       30: // ---- ukonceni handshake: shodit Execute, pockat az kamera shodi stav ----
           "COG_ETIKETA_is3800-ExecuteCommand/JobLoad" := FALSE;
           IF NOT "COG_ETIKETA_is3800-CommandCompleted"
               AND NOT "COG_ETIKETA_is3800-CommandFailed" THEN
               #Kam_Etiketa_Job.krok := 0;
           END_IF;

       ELSE
           #Kam_Etiketa_Job.krok := 0;
   END_CASE;

   // casovac timeoutu bezi v krocich 10..30
   #TIMER.TIMER_3.TON(IN := #Kam_Etiketa_Job.krok >= 10,
                      PT := #Kam_Etiketa_Job.timeout);
   IF #TIMER.TIMER_3.Q AND #Kam_Etiketa_Job.krok = 30 THEN
       #Kam_Etiketa_Job.krok := 0;                         // pojistka, kdyby kamera stav neshodila
   END_IF;

   #Kam_Etiketa_Job.odesli_pamet := "DB_HMI_recype".ODESLI_dATA;

   // kontrola: v klidu musi job v kamere odpovidat recepture
   #Kam_Etiketa_Job.nesouhlasi := #Kam_Etiketa_Job.krok = 0
   AND #Kam_Etiketa_Job.pozadovany > 0
   AND "COG_ETIKETA_is3800-Online"
   AND WORD_TO_INT("COG_ETIKETA_is3800-Current Job ID") <> #Kam_Etiketa_Job.pozadovany;
END_REGION

REGION Network 23: EXTERNAL_TRIGER
   RUNG wire#powerrail
      { S7_Templates := "SrcType := Int" } EQ_Contact(in1 := #SQCR, in2 := #STEP_5_HOME)
      Contact( "INICIALIZACE_RUN" )
      I_Contact( #TRIG.inicial_ok_op )
      Contact( "AUTOMAT" )
      S_Coil( #HMI.reset_fronty )
      S_Coil( #TRIG.inicial_ok_op )
   END_RUNG
   RUNG wire#powerrail
      Contact( "FirstScan" )
      S_Coil( #HMI.reset_fronty )
      Move(in := 0, out1 => "DB_HMI_recype".obsazenost_fronty, out2 => #zpracovani_dat[1].balik_den)
   END_RUNG
   // the same network as SCL:
   IF (#SQCR = #STEP_5_HOME) AND "INICIALIZACE_RUN" AND NOT #TRIG.inicial_ok_op AND "AUTOMAT" THEN
       #HMI.reset_fronty := TRUE;
       #TRIG.inicial_ok_op := TRUE;
   END_IF;
   IF "FirstScan" THEN
       #HMI.reset_fronty := TRUE;
       "DB_HMI_recype".obsazenost_fronty := 0;
       #zpracovani_dat[1].balik_den := 0;
   END_IF;
END_REGION

REGION Network 24: ETERNAL_TRIGR_INICIAL
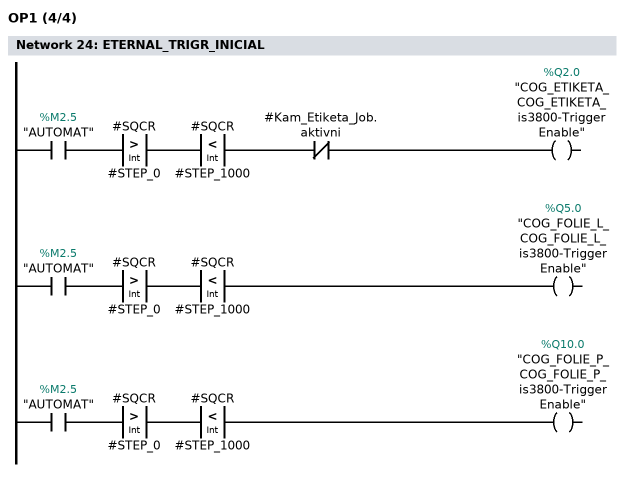
   RUNG wire#powerrail
      Contact( "AUTOMAT" )
      { S7_Templates := "SrcType := Int" } GT_Contact(in1 := #SQCR, in2 := #STEP_0)
      { S7_Templates := "SrcType := Int" } LT_Contact(in1 := #SQCR, in2 := #STEP_1000)
      I_Contact( #Kam_Etiketa_Job.aktivni )
      Coil( "COG_ETIKETA_COG_ETIKETA_is3800-TriggerEnable" )
   END_RUNG
   RUNG wire#powerrail
      Contact( "AUTOMAT" )
      { S7_Templates := "SrcType := Int" } GT_Contact(in1 := #SQCR, in2 := #STEP_0)
      { S7_Templates := "SrcType := Int" } LT_Contact(in1 := #SQCR, in2 := #STEP_1000)
      Coil( "COG_FOLIE_L_COG_FOLIE_L_is3800-TriggerEnable" )
   END_RUNG
   RUNG wire#powerrail
      Contact( "AUTOMAT" )
      { S7_Templates := "SrcType := Int" } GT_Contact(in1 := #SQCR, in2 := #STEP_0)
      { S7_Templates := "SrcType := Int" } LT_Contact(in1 := #SQCR, in2 := #STEP_1000)
      Coil( "COG_FOLIE_P_COG_FOLIE_P_is3800-TriggerEnable" )
   END_RUNG
   // the same network as SCL:
   "COG_ETIKETA_COG_ETIKETA_is3800-TriggerEnable" := "AUTOMAT" AND (#SQCR > #STEP_0) AND (#SQCR < #STEP_1000) AND NOT #Kam_Etiketa_Job.aktivni;
   "COG_FOLIE_L_COG_FOLIE_L_is3800-TriggerEnable" := "AUTOMAT" AND (#SQCR > #STEP_0) AND (#SQCR < #STEP_1000);
   "COG_FOLIE_P_COG_FOLIE_P_is3800-TriggerEnable" := "AUTOMAT" AND (#SQCR > #STEP_0) AND (#SQCR < #STEP_1000);
END_REGION

REGION Network 25: hmi
END_REGION

REGION Network 26 (SCL): VYRAZENI MANUAL
   (* #Test_tp_ka12(IN := "DB_Manual".test_vyr,
                 PT := T#500MS);

   "-KA12" := #Test_tp_ka12.Q;

   // testovací bit se sám shodí → každý Modify TRUE = jeden pulz
   IF "DB_Manual".test_vyr THEN
       "DB_Manual".test_vyr := FALSE;
   END_IF; *)
END_REGION
END_FUNCTION_BLOCK

FUNCTION_BLOCK "FB_CamManual"
{ S7_Optimized_Access := 'TRUE' }
VERSION : 0.1
   VAR_INPUT 
      xManEtiketa : Bool;   // ruční test etiketa
      xManFolie : Bool;   // ruční test folie
      tLightDelay : Time := T#100ms;   // náběh světel
      tTrigPulse : Time := T#50ms;   // d0lka triggeru
   END_VAR

   VAR 
      tonEt {InstructionName := 'TON_TIME'; LibVersion := '1.0'; S7_SetPoint := 'False'} : TON_TIME;
      tpEt {InstructionName := 'TP_TIME'; LibVersion := '1.0'} : TP_TIME;
      tonFo {InstructionName := 'TON_TIME'; LibVersion := '1.0'} : TON_TIME;
      tpFo {InstructionName := 'TP_TIME'; LibVersion := '1.0'} : TP_TIME;
   END_VAR


BEGIN
	// ---------- ETIKETA ----------
	#tonEt(IN := #xManEtiketa,
	       PT := #tLightDelay);
	#tpEt(IN := #tonEt.Q,
	      PT := #tTrigPulse);
	
	IF #xManEtiketa THEN
	    "-KA1" := TRUE;
	    "-KA2" := TRUE;
	END_IF;
	IF #tpEt.Q THEN
	    "COG_ETIKETA_COG_ETIKETA_is3800-Trigger" := TRUE;
	END_IF;
	
	// ---------- FÓLIE ----------
	#tonFo(IN := #xManFolie,
	       PT := #tLightDelay);
	#tpFo(IN := #tonFo.Q,
	      PT := #tTrigPulse);
	
	IF #xManFolie THEN
	    "-KA3" := TRUE;
	    "-KA4" := TRUE;
	    "-KA5" := TRUE;
	END_IF;
	IF #tpFo.Q THEN
	    "COG_FOLIE_L_is3800-Trigger" := TRUE;
	    "COG_FOLIE_P_is3800-Trigger" := TRUE;
	END_IF;
END_FUNCTION_BLOCK

FUNCTION_BLOCK "OP2"   // FB51, LAD
{ S7_Optimized_Access := 'FALSE' }
// stored: AutoNumber false, SetENOAutomatically false
   VAR
      CONTROL_MAN : Struct
         B0 : Bool;
         B1 : Bool;
         B2 : Bool;
         B3 : Bool;
         B4 : Bool;
         B5 : Bool;
         B6 : Bool;
         B7 : Bool;
         B8 : Bool;
         B9 : Bool;
         odfuk_1 : Bool;
         odfuk_2 : Bool;
         B12 : Bool;
         B13 : Bool;
         B14 : Bool;
         B15 : Bool;
         B16 : Bool;
         B17 : Bool;
         B18 : Bool;
         B19 : Bool;
         B20 : Bool;
         B21 : Bool;
         B22 : Bool;
         B23 : Bool;
         B24 : Bool;
         B25 : Bool;
         B26 : Bool;
         B27 : Bool;
         B28 : Bool;
         B29 : Bool;
         B30 : Bool;
         B31 : Bool;
      END_STRUCT;
      CONTROL_AUTOMAT : Struct
         connect : Bool;
         send : Bool;
         reciv : Bool;
         trcv : Bool;
         discon : Bool;
         B5 : Bool;
         B6 : Bool;
         B7 : Bool;
         B8 : Bool;
         B9 : Bool;
         B10 : Bool;
         B11 : Bool;
         B12 : Bool;
         B13 : Bool;
         B14 : Bool;
         B15 : Bool;
         B16 : Bool;
         B17 : Bool;
         B18 : Bool;
         B19 : Bool;
         B20 : Bool;
         B21 : Bool;
         B22 : Bool;
         B23 : Bool;
         B24 : Bool;
         B25 : Bool;
         B26 : Bool;
         B27 : Bool;
         B28 : Bool;
         B29 : Bool;
         B30 : Bool;
         B31 : Bool;
      END_STRUCT;
      SENSORS : Struct
         S0 : Bool;
         S1 : Bool;
         S2 : Bool;
         S3 : Bool;
         S4 : Bool;
         S5 : Bool;
         S6 : Bool;
         S7 : Bool;
         S8 : Bool;   // KARUSEL JE NATOČEN PŘÍPRAVKEM A K BRÁNĚ
         S9 : Bool;
         S10 : Bool;
         S11 : Bool;
         S12 : Bool;
         S13 : Bool;
         S14 : Bool;
         S15 : Bool;
         S16 : Bool;
         S17 : Bool;
         S18 : Bool;
         S19 : Bool;
         S20 : Bool;
         S21 : Bool;
         S22 : Bool;
         S23 : Bool;
         S24 : Bool;
         S25 : Bool;
         S26 : Bool;
         S27 : Bool;
         S28 : Bool;
         S29 : Bool;
         S30 : Bool;
         S31 : Bool;
      END_STRUCT;
      SENSORS_1 : Struct
         S0 : Bool;
         S1 : Bool;
         S2 : Bool;
         S3 : Bool;
         S4 : Bool;
         S5 : Bool;
         S6 : Bool;
         S7 : Bool;
         S8 : Bool;
         S9 : Bool;
         S10 : Bool;
         S11 : Bool;
         S12 : Bool;
         S13 : Bool;
         S14 : Bool;
         S15 : Bool;
         S16 : Bool;
         S17 : Bool;
         S18 : Bool;
         S19 : Bool;
         S20 : Bool;
         S21 : Bool;
         S22 : Bool;
         S23 : Bool;
         S24 : Bool;
         S25 : Bool;
         S26 : Bool;
         S27 : Bool;
         S28 : Bool;
         S29 : Bool;
         S30 : Bool;
         S31 : Bool;
      END_STRUCT;
      S_0 : "SENSOR";
      S_1 : "SENSOR";
      S_2 { S7_SetPoint := 'True'} : "SENSOR";
      S_3 { S7_SetPoint := 'True'} : "SENSOR";
      S_4 { S7_SetPoint := 'True'} : "SENSOR";
      S_5 { S7_SetPoint := 'True'} : "SENSOR";
      S_6 { S7_SetPoint := 'True'} : "SENSOR";
      S_7 { S7_SetPoint := 'True'} : "SENSOR";
      S_8 { S7_SetPoint := 'True'} : "SENSOR";
      S_9 { S7_SetPoint := 'True'} : "SENSOR";
      S_10 { S7_SetPoint := 'True'} : "SENSOR";
      S_11 { S7_SetPoint := 'True'} : "SENSOR";
      S_12 { S7_SetPoint := 'True'} : "SENSOR";
      S_13 { S7_SetPoint := 'True'} : "SENSOR";
      S_14 { S7_SetPoint := 'True'} : "SENSOR";
      S_15 { S7_SetPoint := 'True'} : "SENSOR";
      S_16 { S7_SetPoint := 'True'} : "SENSOR";
      M_1 : "MOTOR_CONTROL_BLOCK";
      M_2 { S7_SetPoint := 'True'} : "MOTOR_CONTROL_BLOCK";
      M_3 { S7_SetPoint := 'True'} : "MOTOR_CONTROL_BLOCK";
      SQCR { S7_SetPoint := 'True'} : Int;
      hmi_sqcr : Int;
      TRIG : Struct
         inicial_ok_op : Bool;
         T2 : Bool;
         T3 : Bool;
         T4 : Bool;
         T5 : Bool;
         T6 : Bool;
         T7 : Bool;
         T8 : Bool;
         T9 : Bool;
         T10 : Bool;
         T11 : Bool;
         T12 : Bool;
         T13 : Bool;
         T14 : Bool;
         T15 : Bool;
         T16 : Bool;
         op_1_ready : Bool;
      END_STRUCT;
      MEMOR : Struct
         n_trig_vypnuti : Bool;
         M1 : Bool;
         M2 : Bool;
         M3 : Bool;
         M4 : Bool;
         p_trig_odavacka : Bool;
         M6 : Bool;
         M7 : Bool;
         M8 : Bool;
         M9 : Bool;
         M10 : Bool;
         M11 : Bool;
         RESET_ERROR : Bool;
         M13 : Bool;
         M14 : Bool;
         M15 : Bool;
         SETOVANI_START : Bool;
         M17 : Bool;
         M18 : Bool;
         M19 : Bool;
         M20 : Bool;
         M21 : Bool;
         M22 : Bool;
         M23 : Bool;
         M24 : Bool;
         M25 : Bool;
         M26 : Bool;
         M27 : Bool;
         M28 : Bool;
         M29 : Bool;
         M30 : Bool;
         N_TRIG_SAFETY : Bool;
         M32 : Bool;
         M33 : Bool;
         start_caklu : Bool;
         M35 : Bool;
         M36 : Bool;
         M37 : Bool;
         M38 : Bool;
         M39 : Bool;
         ALARM_GLOBAL : Bool;
         M41 : Bool;
         M42 : Bool;
         M43 : Bool;
         M44 : Bool;
         M45 : Bool;
         M46 : Bool;
         M47 : Bool;
         M48 : Bool;
         M49 : Bool;
         wrong_p_trig : Bool;
         alarm_p_trig : Bool;
         M52 : Bool;
         M53 : Bool;
         M54 : Bool;
         M55 : Bool;
         M56 : Bool;
         M57 : Bool;
         M58 : Bool;
         M59 : Bool;
         M60 : Bool;
         M61 : Bool;
         M62 : Bool;
         M63 : Bool;
      END_STRUCT;
      "TIMER" : Struct
         TIMER_0 : IEC_TIMER;
         TIMER_1 : IEC_TIMER;
         TIMER_2 : IEC_TIMER;
         TIMER_3 : IEC_TIMER;
         TIMER_4 : IEC_TIMER;
         air : IEC_TIMER;
         TIMER_6 : IEC_TIMER;
         TIMER_7 : IEC_TIMER;
      END_STRUCT;
      HMI : Struct
         povoleni_volby_receptu : Bool;
         "svetlo_on/off" : Bool;
         ALARM_VIDITELNOST : Bool;
         hmi_3 : Bool;
         hmi_4 : Bool;
         hmi_5 : Bool;
         hmi_6 : Bool;
         hmi_7 : Bool;
         hmi_8 : Bool;
         hmi_9 : Bool;
         hmi_10 : Bool;
         hmi_11 : Bool;
         hmi_12 : Bool;
         hmi_13 : Bool;
         hmi_14 : Bool;
         hmi_15 : Bool;
      END_STRUCT;
      int_hodnota_zpravy { ExternalAccessible := 'False'; ExternalVisible := 'False'; ExternalWritable := 'False'} : Word;
      array_do_db AT int_hodnota_zpravy : Array[1..2] of Byte;
      CTRV_LEN { ExternalAccessible := 'False'; ExternalVisible := 'False'; ExternalWritable := 'False'} : UDInt;
      TCON_Instance { S7_SetPoint := 'True'} : TCON;
      TSEND_Instance { S7_SetPoint := 'True'} : TSEND;
      TRCV_Instance { S7_SetPoint := 'True'} : TRCV;
      TDISCON_Instance { S7_SetPoint := 'True'} : TDISCON;
      Tisk : Struct
         pole2_index_bajt : Int := 14;   // bajt rámce s číslem proměnné
         pole2_index_hodnota : Byte := 16#1;   // číslo proměnné pole 2 (pole 1 = 0)
         datum_chyba : Bool;   // datum přepsáno na XX.XX.XXXX
         pole2_kratky : Bool := true;
         jeden_ramec : Bool;
      END_STRUCT;
   END_VAR
   VAR_TEMP
      DATA : Array[0..255] of Char;
      ARRAY_NULL : Array[1..8] of Bool;
      ARRAY_PRAZDNE : Array[0..255] of Byte;
      j : Int;
      L1 : Int;
      p : Int;
   END_VAR
   VAR CONSTANT
      STEP_0 : Int := 0;
      step_2 : Int := 2;
      STEP_4 : Int := 4;
      STEP_5_HOME : Int := 5;
      STEP_7 : Int := 7;
      STEP_10 : Int := 10;
      STEP_15 : Int := 15;
      STEP_20 : Int := 20;
      STEP_23 : Int := 23;
      STEP_25 : Int := 25;
      STEP_27 : Int := 27;
      STEP_30 : Int := 30;
      STEP_35 : Int := 35;
      STEP_37 : Int := 37;
      STEP_40 : Int := 40;
      STEP_43 : Int := 43;
      STEP_45 : Int := 45;
      STEP_50 : Int := 50;
      STEP_55 : Int := 55;
      STEP_60 : Int := 60;
      STEP_65 : Int := 65;
      STEP_70 : Int := 70;
      STEP_73 : Int := 73;
      STEP_75 : Int := 75;
      STEP_80 : Int := 80;
      STEP_83 : Int := 83;
      STEP_85 : Int := 85;
      STEP_90 : Int := 90;
      STEP_93 : Int := 93;
      STEP_95 : Int := 95;
      STEP_100 : Int := 100;
      STEP_105 : Int := 105;
      STEP_110 : Int := 110;
      STEP_113 : Int := 113;
      STEP_115 : Int := 115;
      STEP_120 : Int := 120;
      STEP_125 : Int := 125;
      STEP_130 : Int := 130;
      STEP_135 : Int := 135;
      STEP_140 : Int := 140;
      STEP_145 : Int := 145;
      STEP_150 : Int := 150;
      STEP_155 : Int := 155;
      STEP_1000 : Int := 1000;
      STEP_1001 : Int := 1001;
      STEP_1002 : Int := 1002;
      STEP_1003 : Int := 1003;
      STEP_1004 : Int := 1004;
      STEP_1005 : Int := 1005;
      STEP_1010 : Int := 1010;
      STEP_1015 : Int := 1015;
      STEP_1020 : Int := 1020;
      STEP_1025 : Int := 1025;
      STEP_3000 : Int := 3000;
      STEP_3005 : Int := 3005;
      STEP_3010 : Int := 3010;
      STEP_3015 : Int := 3015;
      STEP_3020 : Int := 3020;
      STEP_2000 : Int := 2000;
      string_null : String;
      char_null : Char;
      text_kartacek : String := 'Kartacek';
      string_kar_A : String := 'A';
      string_kar_B : String := 'B';
   END_VAR
   VAR_TEMP   // added for the SCL form of the ladder/FBD networks
      _w1 : Bool;
      _w2 : Bool;
      _w3 : Bool;
   END_VAR
BEGIN

REGION Network 1: manuali ovladani reset
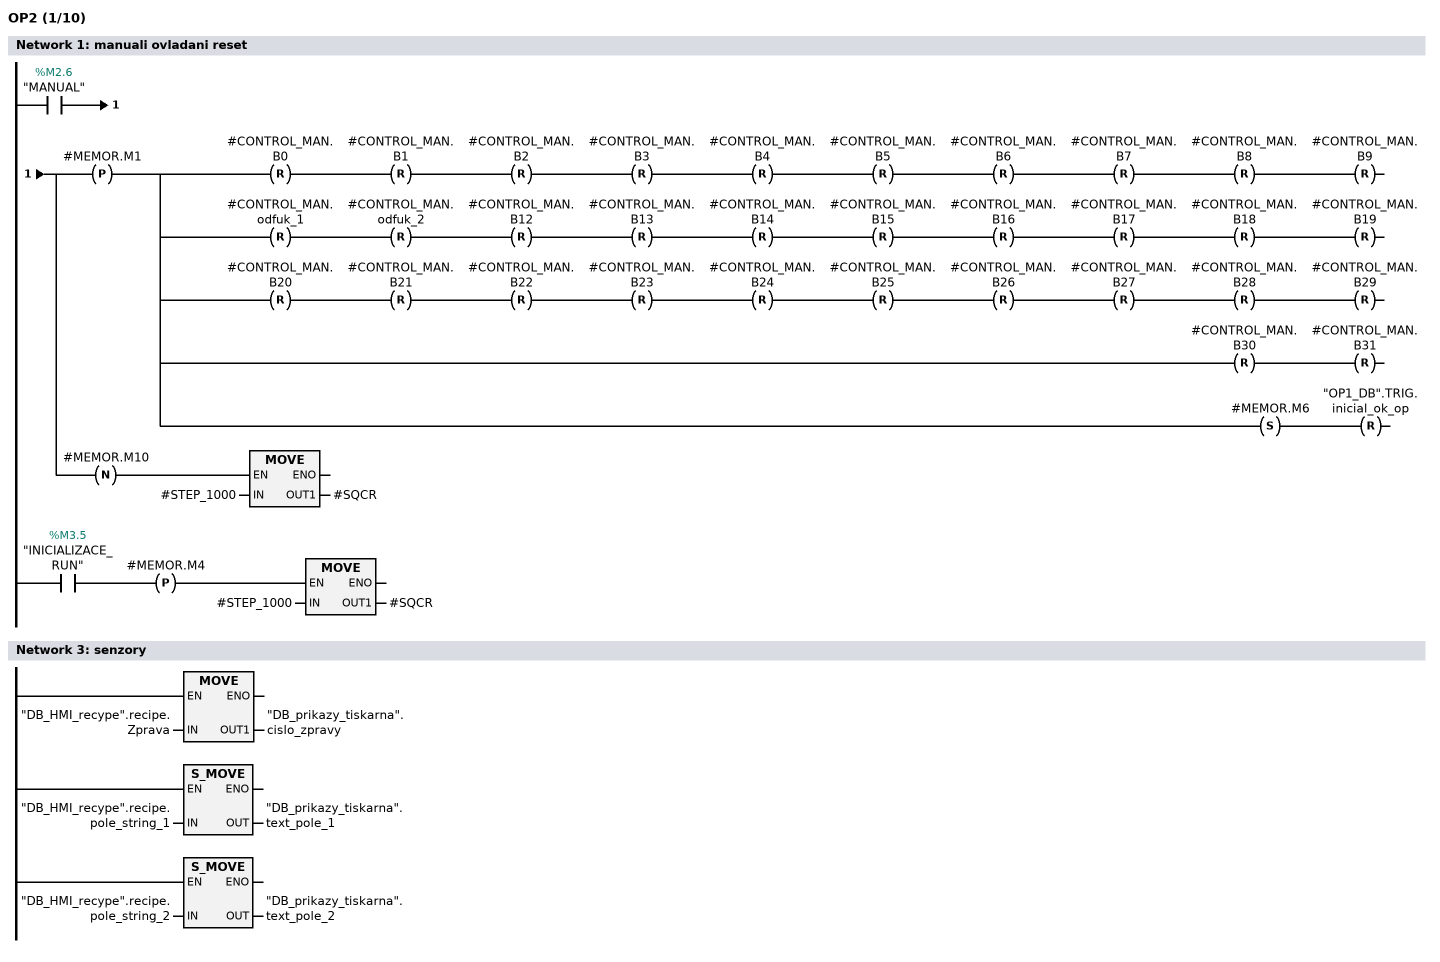
   RUNG wire#powerrail
      Contact( "MANUAL" )
      wire#w1
      P_Trig( #MEMOR.M1 )
      wire#w2
      R_Coil( #CONTROL_MAN.B0 )
      R_Coil( #CONTROL_MAN.B1 )
      R_Coil( #CONTROL_MAN.B2 )
      R_Coil( #CONTROL_MAN.B3 )
      R_Coil( #CONTROL_MAN.B4 )
      R_Coil( #CONTROL_MAN.B5 )
      R_Coil( #CONTROL_MAN.B6 )
      R_Coil( #CONTROL_MAN.B7 )
      R_Coil( #CONTROL_MAN.B8 )
      R_Coil( #CONTROL_MAN.B9 )
   END_RUNG
   RUNG wire#w2
      R_Coil( #CONTROL_MAN.odfuk_1 )
      R_Coil( #CONTROL_MAN.odfuk_2 )
      R_Coil( #CONTROL_MAN.B12 )
      R_Coil( #CONTROL_MAN.B13 )
      R_Coil( #CONTROL_MAN.B14 )
      R_Coil( #CONTROL_MAN.B15 )
      R_Coil( #CONTROL_MAN.B16 )
      R_Coil( #CONTROL_MAN.B17 )
      R_Coil( #CONTROL_MAN.B18 )
      R_Coil( #CONTROL_MAN.B19 )
   END_RUNG
   RUNG wire#w2
      R_Coil( #CONTROL_MAN.B20 )
      R_Coil( #CONTROL_MAN.B21 )
      R_Coil( #CONTROL_MAN.B22 )
      R_Coil( #CONTROL_MAN.B23 )
      R_Coil( #CONTROL_MAN.B24 )
      R_Coil( #CONTROL_MAN.B25 )
      R_Coil( #CONTROL_MAN.B26 )
      R_Coil( #CONTROL_MAN.B27 )
      R_Coil( #CONTROL_MAN.B28 )
      R_Coil( #CONTROL_MAN.B29 )
   END_RUNG
   RUNG wire#w2
      R_Coil( #CONTROL_MAN.B30 )
      R_Coil( #CONTROL_MAN.B31 )
   END_RUNG
   RUNG wire#w2
      S_Coil( #MEMOR.M6 )
      R_Coil( "OP1_DB".TRIG.inicial_ok_op )
   END_RUNG
   RUNG wire#w1
      N_Trig( #MEMOR.M10 )
      Move(in := #STEP_1000, out1 => #SQCR)
   END_RUNG
   RUNG wire#powerrail
      Contact( "INICIALIZACE_RUN" )
      P_Trig( #MEMOR.M4 )
      Move(in := #STEP_1000, out1 => #SQCR)
   END_RUNG
   // the same network as SCL:
   #_w1 := "MANUAL" AND NOT #MEMOR.M1;   // rising edge
   #MEMOR.M1 := "MANUAL";
   IF #_w1 THEN
       #CONTROL_MAN.B0 := FALSE;
       #CONTROL_MAN.B1 := FALSE;
       #CONTROL_MAN.B2 := FALSE;
       #CONTROL_MAN.B3 := FALSE;
       #CONTROL_MAN.B4 := FALSE;
       #CONTROL_MAN.B5 := FALSE;
       #CONTROL_MAN.B6 := FALSE;
       #CONTROL_MAN.B7 := FALSE;
       #CONTROL_MAN.B8 := FALSE;
       #CONTROL_MAN.B9 := FALSE;
       #CONTROL_MAN.odfuk_1 := FALSE;
       #CONTROL_MAN.odfuk_2 := FALSE;
       #CONTROL_MAN.B12 := FALSE;
       #CONTROL_MAN.B13 := FALSE;
       #CONTROL_MAN.B14 := FALSE;
       #CONTROL_MAN.B15 := FALSE;
       #CONTROL_MAN.B16 := FALSE;
       #CONTROL_MAN.B17 := FALSE;
       #CONTROL_MAN.B18 := FALSE;
       #CONTROL_MAN.B19 := FALSE;
       #CONTROL_MAN.B20 := FALSE;
       #CONTROL_MAN.B21 := FALSE;
       #CONTROL_MAN.B22 := FALSE;
       #CONTROL_MAN.B23 := FALSE;
       #CONTROL_MAN.B24 := FALSE;
       #CONTROL_MAN.B25 := FALSE;
       #CONTROL_MAN.B26 := FALSE;
       #CONTROL_MAN.B27 := FALSE;
       #CONTROL_MAN.B28 := FALSE;
       #CONTROL_MAN.B29 := FALSE;
       #CONTROL_MAN.B30 := FALSE;
       #CONTROL_MAN.B31 := FALSE;
       #MEMOR.M6 := TRUE;
       "OP1_DB".TRIG.inicial_ok_op := FALSE;
   END_IF;
   #_w2 := NOT "MANUAL" AND #MEMOR.M10;   // falling edge
   #MEMOR.M10 := "MANUAL";
   IF #_w2 THEN #SQCR := #STEP_1000; END_IF;
   #_w3 := "INICIALIZACE_RUN" AND NOT #MEMOR.M4;   // rising edge
   #MEMOR.M4 := "INICIALIZACE_RUN";
   IF #_w3 THEN #SQCR := #STEP_1000; END_IF;
END_REGION

REGION Network 2: alarmy
END_REGION

REGION Network 3: senzory
   RUNG wire#powerrail
      Move(in := "DB_HMI_recype".recipe.Zprava, out1 => "DB_prikazy_tiskarna".cislo_zpravy)
   END_RUNG
   RUNG wire#powerrail
      S_Move(in := "DB_HMI_recype".recipe.pole_string_1, out => "DB_prikazy_tiskarna".text_pole_1)
   END_RUNG
   RUNG wire#powerrail
      S_Move(in := "DB_HMI_recype".recipe.pole_string_2, out => "DB_prikazy_tiskarna".text_pole_2)
   END_RUNG
   // the same network as SCL:
   "DB_prikazy_tiskarna".cislo_zpravy := "DB_HMI_recype".recipe.Zprava;
   "DB_prikazy_tiskarna".text_pole_1 := "DB_HMI_recype".recipe.pole_string_1;
   "DB_prikazy_tiskarna".text_pole_2 := "DB_HMI_recype".recipe.pole_string_2;
END_REGION

REGION Network 4 (SCL): tiskarna_zpracovani_dat


   #int_hodnota_zpravy := "DB_prikazy_tiskarna".cislo_zpravy;


   //"DB_prikazy_tiskarna".byte_2 := INT_TO_CHAR( "DB_prikazy_tiskarna".cislo_zpravy);
   "DB_prikazy_tiskarna".byte_1 := #array_do_db[1] + 48;
   "DB_prikazy_tiskarna".byte_2 := #array_do_db[2] + 48;


   "DB_prikazy_tiskarna".task[3, 26] := "DB_prikazy_tiskarna".byte_1;
   "DB_prikazy_tiskarna".task[3, 27] := "DB_prikazy_tiskarna".byte_2;











   "DB_prikazy_tiskarna".task[4, 17] := "DB_prikazy_tiskarna".text_pole_1[1];
   "DB_prikazy_tiskarna".task[4, 18] := "DB_prikazy_tiskarna".text_pole_1[2];
   "DB_prikazy_tiskarna".task[4, 19] := "DB_prikazy_tiskarna".text_pole_1[3];
   "DB_prikazy_tiskarna".task[4, 20] := "DB_prikazy_tiskarna".text_pole_1[4];
   "DB_prikazy_tiskarna".task[4, 21] := "DB_prikazy_tiskarna".text_pole_1[5];
   "DB_prikazy_tiskarna".task[4, 22] := "DB_prikazy_tiskarna".text_pole_1[6];
   "DB_prikazy_tiskarna".task[4, 23] := "DB_prikazy_tiskarna".text_pole_1[7];
   "DB_prikazy_tiskarna".task[4, 24] := "DB_prikazy_tiskarna".text_pole_1[8];
   "DB_prikazy_tiskarna".task[4, 25] := "DB_prikazy_tiskarna".text_pole_1[9];
   "DB_prikazy_tiskarna".task[4, 26] := "DB_prikazy_tiskarna".text_pole_1[10];
   "DB_prikazy_tiskarna".task[4, 27] := "DB_prikazy_tiskarna".text_pole_1[11];
   "DB_prikazy_tiskarna".task[4, 28] := "DB_prikazy_tiskarna".text_pole_1[12];
   "DB_prikazy_tiskarna".task[4, 29] := "DB_prikazy_tiskarna".text_pole_1[13];
   "DB_prikazy_tiskarna".task[4, 30] := "DB_prikazy_tiskarna".text_pole_1[14];
   "DB_prikazy_tiskarna".task[4, 31] := "DB_prikazy_tiskarna".text_pole_1[15];
   "DB_prikazy_tiskarna".task[4, 32] := "DB_prikazy_tiskarna".text_pole_1[16];
   "DB_prikazy_tiskarna".task[4, 33] := "DB_prikazy_tiskarna".text_pole_1[17];
   "DB_prikazy_tiskarna".task[4, 34] := "DB_prikazy_tiskarna".text_pole_1[18];
   "DB_prikazy_tiskarna".task[4, 35] := "DB_prikazy_tiskarna".text_pole_1[19];
   "DB_prikazy_tiskarna".task[4, 36] := "DB_prikazy_tiskarna".text_pole_1[20];
   "DB_prikazy_tiskarna".task[4, 37] := "DB_prikazy_tiskarna".text_pole_1[21];
   "DB_prikazy_tiskarna".task[4, 38] := "DB_prikazy_tiskarna".text_pole_1[22];
   "DB_prikazy_tiskarna".task[4, 39] := "DB_prikazy_tiskarna".text_pole_1[23];
   "DB_prikazy_tiskarna".task[4, 40] := "DB_prikazy_tiskarna".text_pole_1[24];
   "DB_prikazy_tiskarna".task[4, 41] := "DB_prikazy_tiskarna".text_pole_1[25];
   "DB_prikazy_tiskarna".task[4, 42] := "DB_prikazy_tiskarna".text_pole_1[26];
   "DB_prikazy_tiskarna".task[4, 43] := "DB_prikazy_tiskarna".text_pole_1[27];
   "DB_prikazy_tiskarna".task[4, 44] := "DB_prikazy_tiskarna".text_pole_1[28];
   "DB_prikazy_tiskarna".task[4, 45] := "DB_prikazy_tiskarna".text_pole_1[29];
   "DB_prikazy_tiskarna".task[4, 46] := "DB_prikazy_tiskarna".text_pole_1[30];






   IF "DB_HMI_recype".recipe.pole_string_2[3] <> '.' OR "DB_HMI_recype".recipe.pole_string_2[6] <> '.' THEN
       "DB_HMI_recype".recipe.pole_string_2 := 'XX.XX.XXXX';
   END_IF;



   // ===================== POLE 2 - DATUM SPOTREBY (radek 5) =====================
   // Samostatny ramec CF stejny jako pole 1 (radek 4), lisi se cislem promenne,
   // delkou textu a obsahem. Odesila se v kroku 130 (ADRESACE_POLE = 5).

   // chybne datum (prepsane na XX) -> priznak pro alarm / vyrazeni
   #Tisk.datum_chyba := "DB_HMI_recype".recipe.pole_string_2 = 'XX.XX.XXXX';

   // hlavicka ramce = kopie hlavicky pole 1 (bajty 0..16)
   FOR #j := 0 TO 16 DO
       "DB_prikazy_tiskarna".task[5, #j] := "DB_prikazy_tiskarna".task[4, #j];
   END_FOR;

   // cislo promenne pole 2 - bajt nastavitelny (12/13/14), overit na tiskarne
   IF #Tisk.pole2_index_bajt >= 12 AND #Tisk.pole2_index_bajt <= 14 THEN
       "DB_prikazy_tiskarna".task[5, #Tisk.pole2_index_bajt] := #Tisk.pole2_index_hodnota;
   END_IF;

   // datum - vzdy 10 znaku (DD.MM.RRRR nebo XX.XX.XXXX)
   "DB_prikazy_tiskarna".task[5, 17] := "DB_prikazy_tiskarna".text_pole_2[1];
   "DB_prikazy_tiskarna".task[5, 18] := "DB_prikazy_tiskarna".text_pole_2[2];
   "DB_prikazy_tiskarna".task[5, 19] := "DB_prikazy_tiskarna".text_pole_2[3];
   "DB_prikazy_tiskarna".task[5, 20] := "DB_prikazy_tiskarna".text_pole_2[4];
   "DB_prikazy_tiskarna".task[5, 21] := "DB_prikazy_tiskarna".text_pole_2[5];
   "DB_prikazy_tiskarna".task[5, 22] := "DB_prikazy_tiskarna".text_pole_2[6];
   "DB_prikazy_tiskarna".task[5, 23] := "DB_prikazy_tiskarna".text_pole_2[7];
   "DB_prikazy_tiskarna".task[5, 24] := "DB_prikazy_tiskarna".text_pole_2[8];
   "DB_prikazy_tiskarna".task[5, 25] := "DB_prikazy_tiskarna".text_pole_2[9];
   "DB_prikazy_tiskarna".task[5, 26] := "DB_prikazy_tiskarna".text_pole_2[10];

   IF #Tisk.pole2_kratky THEN
       // --- 10 znaku: upravit delky v hlavicce ---
       "DB_prikazy_tiskarna".task[5, 5] := 16#28;   // delka ramce od bajtu 6 = 40
       "DB_prikazy_tiskarna".task[5, 8] := 16#00;
       "DB_prikazy_tiskarna".task[5, 9] := 16#24;   // delka dat prikazu od bajtu 10 = 36
       "DB_prikazy_tiskarna".task[5, 15] := 16#00;
       "DB_prikazy_tiskarna".task[5, 16] := 16#0A;   // delka textu = 10 znaku
       // za datem 19 x 00 (bajty 27..45), dal nic
       FOR #j := 27 TO 65 DO
           "DB_prikazy_tiskarna".task[5, #j] := 16#00;
       END_FOR;
   ELSE
       // --- 30 znaku (puvodni varianta): delky z hlavicky pole 1, doplnit mezerami ---
       FOR #j := 27 TO 46 DO
           "DB_prikazy_tiskarna".task[5, #j] := 16#20;
       END_FOR;
       FOR #j := 47 TO 65 DO
           "DB_prikazy_tiskarna".task[5, #j] := 16#00;
       END_FOR;
   END_IF;

   // ===== OBE POLE V JEDNOM RAMCI CF: 20 promennych, delka 1 bajt =====
   IF #Tisk.jeden_ramec THEN
       #L1 := LEN("DB_prikazy_tiskarna".text_pole_1);
       IF #L1 > 30 THEN
           #L1 := 30;
       END_IF;

       FOR #j := 15 TO 120 DO
           "DB_prikazy_tiskarna".task[4, #j] := 16#00;
       END_FOR;

       // promenna 1: delka (1 bajt) + Puvod
       "DB_prikazy_tiskarna".task[4, 16] := INT_TO_BYTE(#L1);
       FOR #j := 1 TO #L1 DO
           "DB_prikazy_tiskarna".task[4, 16 + #j] := "DB_prikazy_tiskarna".text_pole_1[#j];
       END_FOR;
       #p := 17 + #L1;

       // promenna 2: delka (1 bajt) + datum
       "DB_prikazy_tiskarna".task[4, #p] := 16#0A;
       FOR #j := 1 TO 10 DO
           "DB_prikazy_tiskarna".task[4, #p + #j] := "DB_prikazy_tiskarna".text_pole_2[#j];
       END_FOR;
       #p := #p + 11;

       // promenne 3..20 prazdne = 18 x 00 (uz vycisteno)
       #p := #p + 18;

       "DB_prikazy_tiskarna".task[4, 4] := 16#00;
       "DB_prikazy_tiskarna".task[4, 5] := INT_TO_BYTE(#p - 6);
       "DB_prikazy_tiskarna".task[4, 8] := 16#00;
       "DB_prikazy_tiskarna".task[4, 9] := INT_TO_BYTE(#p - 10);
   END_IF;
END_REGION

REGION Network 5: příkazy k odeslání z bafru
   // 2 = STOP TISKU
   // 3 = VÝBĚR ZPRÁVY
   // 6 = NASTAVENÍ NEBAFROVÁNÍ A SMAZÁNÍ PŘEDEŠLÍCH DAT
   // 4 = ZAPSÁNÍ DO VARIABILNÍHO POLE 1
   // 5 = ZAPSÁNÍ DO VARIABILNÍHO POLE 2
   // 1 = START TISKU
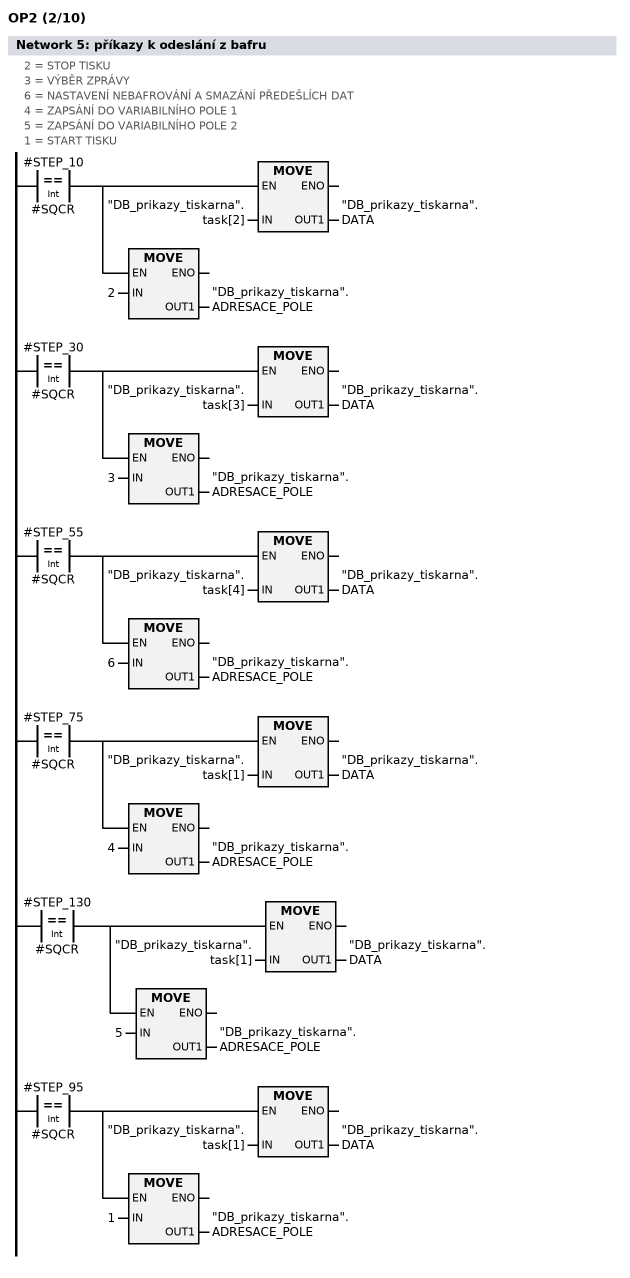
   RUNG wire#powerrail
      { S7_Templates := "SrcType := Int" } EQ_Contact(in1 := #STEP_10, in2 := #SQCR)
      wire#w1
      Move(in := "DB_prikazy_tiskarna".task[2], out1 => "DB_prikazy_tiskarna".DATA)
   END_RUNG
   RUNG wire#w1
      Move(in := 2, out1 => "DB_prikazy_tiskarna".ADRESACE_POLE)
   END_RUNG
   RUNG wire#powerrail
      { S7_Templates := "SrcType := Int" } EQ_Contact(in1 := #STEP_30, in2 := #SQCR)
      wire#w2
      Move(in := "DB_prikazy_tiskarna".task[3], out1 => "DB_prikazy_tiskarna".DATA)
   END_RUNG
   RUNG wire#w2
      Move(in := 3, out1 => "DB_prikazy_tiskarna".ADRESACE_POLE)
   END_RUNG
   RUNG wire#powerrail
      { S7_Templates := "SrcType := Int" } EQ_Contact(in1 := #STEP_55, in2 := #SQCR)
      wire#w3
      Move(in := "DB_prikazy_tiskarna".task[4], out1 => "DB_prikazy_tiskarna".DATA)
   END_RUNG
   RUNG wire#w3
      Move(in := 6, out1 => "DB_prikazy_tiskarna".ADRESACE_POLE)
   END_RUNG
   RUNG wire#powerrail
      { S7_Templates := "SrcType := Int" } EQ_Contact(in1 := #STEP_75, in2 := #SQCR)
      wire#w4
      Move(in := "DB_prikazy_tiskarna".task[1], out1 => "DB_prikazy_tiskarna".DATA)
   END_RUNG
   RUNG wire#w4
      Move(in := 4, out1 => "DB_prikazy_tiskarna".ADRESACE_POLE)
   END_RUNG
   RUNG wire#powerrail
      { S7_Templates := "SrcType := Int" } EQ_Contact(in1 := #STEP_130, in2 := #SQCR)
      wire#w5
      Move(in := "DB_prikazy_tiskarna".task[1], out1 => "DB_prikazy_tiskarna".DATA)
   END_RUNG
   RUNG wire#w5
      Move(in := 5, out1 => "DB_prikazy_tiskarna".ADRESACE_POLE)
   END_RUNG
   RUNG wire#powerrail
      { S7_Templates := "SrcType := Int" } EQ_Contact(in1 := #STEP_95, in2 := #SQCR)
      wire#w6
      Move(in := "DB_prikazy_tiskarna".task[1], out1 => "DB_prikazy_tiskarna".DATA)
   END_RUNG
   RUNG wire#w6
      Move(in := 1, out1 => "DB_prikazy_tiskarna".ADRESACE_POLE)
   END_RUNG
   // the same network as SCL:
   IF #STEP_10 = #SQCR THEN
       "DB_prikazy_tiskarna".DATA := "DB_prikazy_tiskarna".task[2];
       "DB_prikazy_tiskarna".ADRESACE_POLE := 2;
   END_IF;
   IF #STEP_30 = #SQCR THEN
       "DB_prikazy_tiskarna".DATA := "DB_prikazy_tiskarna".task[3];
       "DB_prikazy_tiskarna".ADRESACE_POLE := 3;
   END_IF;
   IF #STEP_55 = #SQCR THEN
       "DB_prikazy_tiskarna".DATA := "DB_prikazy_tiskarna".task[4];
       "DB_prikazy_tiskarna".ADRESACE_POLE := 6;
   END_IF;
   IF #STEP_75 = #SQCR THEN
       "DB_prikazy_tiskarna".DATA := "DB_prikazy_tiskarna".task[1];
       "DB_prikazy_tiskarna".ADRESACE_POLE := 4;
   END_IF;
   IF #STEP_130 = #SQCR THEN
       "DB_prikazy_tiskarna".DATA := "DB_prikazy_tiskarna".task[1];
       "DB_prikazy_tiskarna".ADRESACE_POLE := 5;
   END_IF;
   IF #STEP_95 = #SQCR THEN
       "DB_prikazy_tiskarna".DATA := "DB_prikazy_tiskarna".task[1];
       "DB_prikazy_tiskarna".ADRESACE_POLE := 1;
   END_IF;
END_REGION

REGION Network 6: CONTROL BLOCK tiskarna
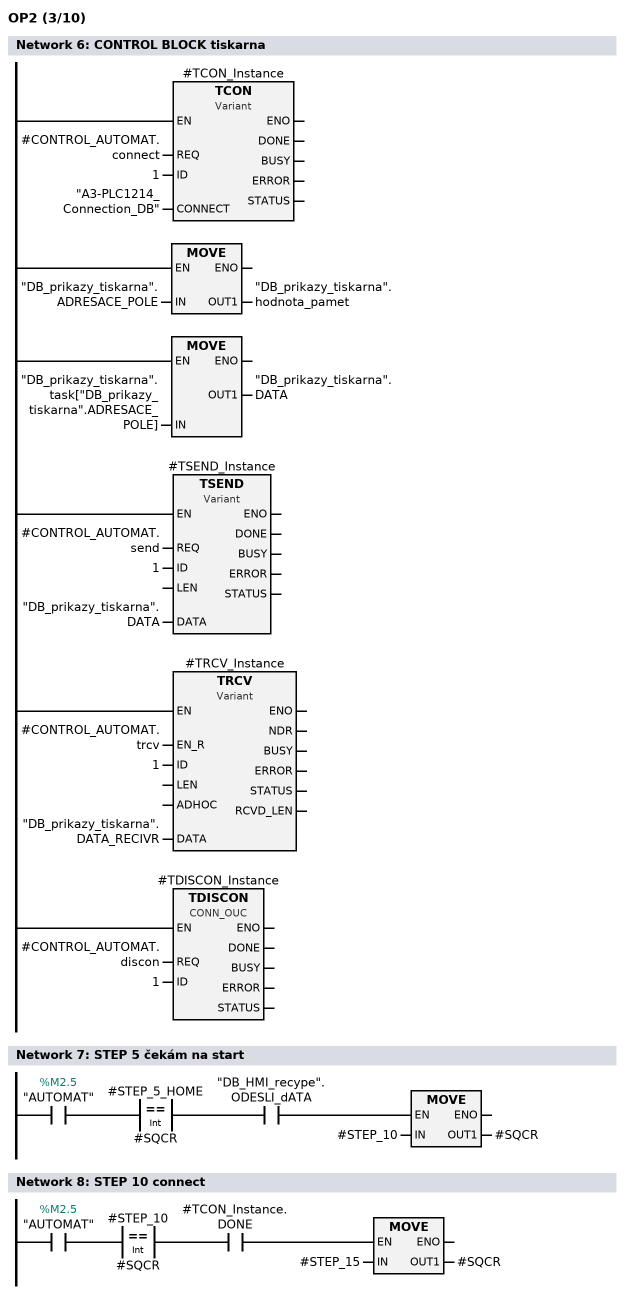
   RUNG wire#powerrail
      { S7_Templates := "[con_type := Variant, id_type := CONN_OUC]" } #TCON_Instance.TCON(REQ := #CONTROL_AUTOMAT.connect, ID := 1, CONNECT := "A3-PLC1214_Connection_DB", DONE =>, BUSY =>, ERROR =>, STATUS =>)
   END_RUNG
   RUNG wire#powerrail
      Move(in := "DB_prikazy_tiskarna".ADRESACE_POLE, out1 => "DB_prikazy_tiskarna".hodnota_pamet)
   END_RUNG
   RUNG wire#powerrail
      Move(in := "DB_prikazy_tiskarna".task["DB_prikazy_tiskarna".ADRESACE_POLE], out1 => "DB_prikazy_tiskarna".DATA)
   END_RUNG
   RUNG wire#powerrail
      { S7_Templates := "[data_type := Variant, len_type := UDInt, id_type := CONN_OUC]" } #TSEND_Instance.TSEND(REQ := #CONTROL_AUTOMAT.send, ID := 1, LEN :=, DATA := "DB_prikazy_tiskarna".DATA, DONE =>, BUSY =>, ERROR =>, STATUS =>)
   END_RUNG
   RUNG wire#powerrail
      { S7_Templates := "[card := 1, ptr_type := Variant, value_type := UDInt, id_type := CONN_OUC]" } #TRCV_Instance.TRCV(EN_R := #CONTROL_AUTOMAT.trcv, ID := 1, LEN :=, ADHOC :=, DATA := "DB_prikazy_tiskarna".DATA_RECIVR, NDR =>, BUSY =>, ERROR =>, STATUS =>, RCVD_LEN =>)
   END_RUNG
   RUNG wire#powerrail
      { S7_Templates := "id_type := CONN_OUC" } #TDISCON_Instance.TDISCON(REQ := #CONTROL_AUTOMAT.discon, ID := 1, DONE =>, BUSY =>, ERROR =>, STATUS =>)
   END_RUNG
   // the same network as SCL:
   #TCON_Instance(REQ := #CONTROL_AUTOMAT.connect, ID := 1, CONNECT := "A3-PLC1214_Connection_DB");   // TCON
   "DB_prikazy_tiskarna".hodnota_pamet := "DB_prikazy_tiskarna".ADRESACE_POLE;
   "DB_prikazy_tiskarna".DATA := "DB_prikazy_tiskarna".task["DB_prikazy_tiskarna".ADRESACE_POLE];
   #TSEND_Instance(REQ := #CONTROL_AUTOMAT.send, ID := 1, DATA := "DB_prikazy_tiskarna".DATA);   // TSEND
   #TRCV_Instance(EN_R := #CONTROL_AUTOMAT.trcv, ID := 1, DATA := "DB_prikazy_tiskarna".DATA_RECIVR);   // TRCV
   #TDISCON_Instance(REQ := #CONTROL_AUTOMAT.discon, ID := 1);   // TDISCON
END_REGION

REGION Network 7: STEP 5 čekám na start
   RUNG wire#powerrail
      Contact( "AUTOMAT" )
      { S7_Templates := "SrcType := Int" } EQ_Contact(in1 := #STEP_5_HOME, in2 := #SQCR)
      Contact( "DB_HMI_recype".ODESLI_dATA )
      Move(in := #STEP_10, out1 => #SQCR)
   END_RUNG
   // the same network as SCL:
   IF "AUTOMAT" AND (#STEP_5_HOME = #SQCR) AND "DB_HMI_recype".ODESLI_dATA THEN #SQCR := #STEP_10; END_IF;
END_REGION

REGION Network 8: STEP 10 connect
   RUNG wire#powerrail
      Contact( "AUTOMAT" )
      { S7_Templates := "SrcType := Int" } EQ_Contact(in1 := #STEP_10, in2 := #SQCR)
      Contact( #TCON_Instance.DONE )
      Move(in := #STEP_15, out1 => #SQCR)
   END_RUNG
   // the same network as SCL:
   IF "AUTOMAT" AND (#STEP_10 = #SQCR) AND #TCON_Instance.DONE THEN #SQCR := #STEP_15; END_IF;
END_REGION

REGION Network 9: STEP 15 tsend STOP_TISKU
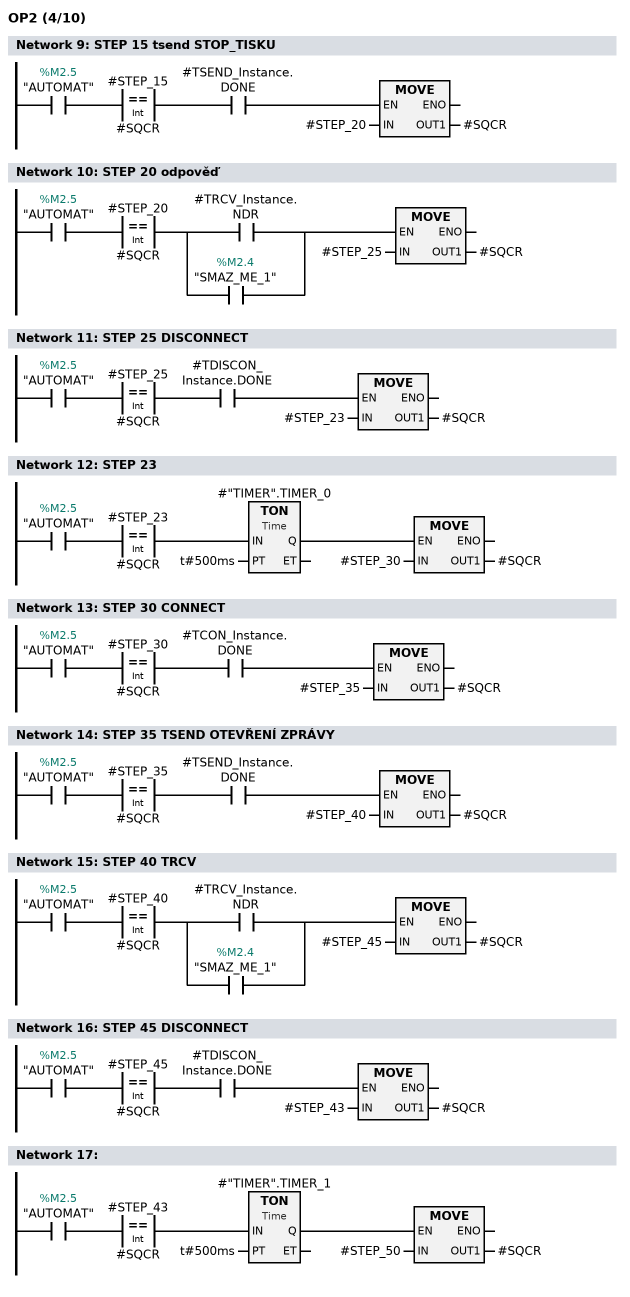
   RUNG wire#powerrail
      Contact( "AUTOMAT" )
      { S7_Templates := "SrcType := Int" } EQ_Contact(in1 := #STEP_15, in2 := #SQCR)
      Contact( #TSEND_Instance.DONE )
      Move(in := #STEP_20, out1 => #SQCR)
   END_RUNG
   // the same network as SCL:
   IF "AUTOMAT" AND (#STEP_15 = #SQCR) AND #TSEND_Instance.DONE THEN #SQCR := #STEP_20; END_IF;
END_REGION

REGION Network 10: STEP 20 odpověď
   RUNG wire#powerrail
      Contact( "AUTOMAT" )
      { S7_Templates := "SrcType := Int" } EQ_Contact(in1 := #STEP_20, in2 := #SQCR)
      wire#w1
      Contact( #TRCV_Instance.NDR )
      wire#w2
      Move(in := #STEP_25, out1 => #SQCR)
   END_RUNG
   RUNG wire#w1
      Contact( "SMAZ_ME_1" )
   END_RUNG wire#w2
   // the same network as SCL:
   IF "AUTOMAT" AND (#STEP_20 = #SQCR) AND (#TRCV_Instance.NDR OR "SMAZ_ME_1") THEN
       #SQCR := #STEP_25;
   END_IF;
END_REGION

REGION Network 11: STEP 25 DISCONNECT
   RUNG wire#powerrail
      Contact( "AUTOMAT" )
      { S7_Templates := "SrcType := Int" } EQ_Contact(in1 := #STEP_25, in2 := #SQCR)
      Contact( #TDISCON_Instance.DONE )
      Move(in := #STEP_23, out1 => #SQCR)
   END_RUNG
   // the same network as SCL:
   IF "AUTOMAT" AND (#STEP_25 = #SQCR) AND #TDISCON_Instance.DONE THEN #SQCR := #STEP_23; END_IF;
END_REGION

REGION Network 12: STEP 23
   RUNG wire#powerrail
      Contact( "AUTOMAT" )
      { S7_Templates := "SrcType := Int" } EQ_Contact(in1 := #STEP_23, in2 := #SQCR)
      { S7_Templates := "time_type := Time" } #"TIMER".TIMER_0.TON(pt := t#500ms, et =>)
      Move(in := #STEP_30, out1 => #SQCR)
   END_RUNG
   // the same network as SCL:
   #"TIMER".TIMER_0.TON(IN := "AUTOMAT" AND (#STEP_23 = #SQCR), PT := t#500ms);
   IF #"TIMER".TIMER_0.Q THEN #SQCR := #STEP_30; END_IF;
END_REGION

REGION Network 13: STEP 30 CONNECT
   RUNG wire#powerrail
      Contact( "AUTOMAT" )
      { S7_Templates := "SrcType := Int" } EQ_Contact(in1 := #STEP_30, in2 := #SQCR)
      Contact( #TCON_Instance.DONE )
      Move(in := #STEP_35, out1 => #SQCR)
   END_RUNG
   // the same network as SCL:
   IF "AUTOMAT" AND (#STEP_30 = #SQCR) AND #TCON_Instance.DONE THEN #SQCR := #STEP_35; END_IF;
END_REGION

REGION Network 14: STEP 35 TSEND OTEVŘENÍ ZPRÁVY
   RUNG wire#powerrail
      Contact( "AUTOMAT" )
      { S7_Templates := "SrcType := Int" } EQ_Contact(in1 := #STEP_35, in2 := #SQCR)
      Contact( #TSEND_Instance.DONE )
      Move(in := #STEP_40, out1 => #SQCR)
   END_RUNG
   // the same network as SCL:
   IF "AUTOMAT" AND (#STEP_35 = #SQCR) AND #TSEND_Instance.DONE THEN #SQCR := #STEP_40; END_IF;
END_REGION

REGION Network 15: STEP 40 TRCV
   RUNG wire#powerrail
      Contact( "AUTOMAT" )
      { S7_Templates := "SrcType := Int" } EQ_Contact(in1 := #STEP_40, in2 := #SQCR)
      wire#w1
      Contact( #TRCV_Instance.NDR )
      wire#w2
      Move(in := #STEP_45, out1 => #SQCR)
   END_RUNG
   RUNG wire#w1
      Contact( "SMAZ_ME_1" )
   END_RUNG wire#w2
   // the same network as SCL:
   IF "AUTOMAT" AND (#STEP_40 = #SQCR) AND (#TRCV_Instance.NDR OR "SMAZ_ME_1") THEN
       #SQCR := #STEP_45;
   END_IF;
END_REGION

REGION Network 16: STEP 45 DISCONNECT
   RUNG wire#powerrail
      Contact( "AUTOMAT" )
      { S7_Templates := "SrcType := Int" } EQ_Contact(in1 := #STEP_45, in2 := #SQCR)
      Contact( #TDISCON_Instance.DONE )
      Move(in := #STEP_43, out1 => #SQCR)
   END_RUNG
   // the same network as SCL:
   IF "AUTOMAT" AND (#STEP_45 = #SQCR) AND #TDISCON_Instance.DONE THEN #SQCR := #STEP_43; END_IF;
END_REGION

REGION Network 17
   RUNG wire#powerrail
      Contact( "AUTOMAT" )
      { S7_Templates := "SrcType := Int" } EQ_Contact(in1 := #STEP_43, in2 := #SQCR)
      { S7_Templates := "time_type := Time" } #"TIMER".TIMER_1.TON(pt := t#500ms, et =>)
      Move(in := #STEP_50, out1 => #SQCR)
   END_RUNG
   // the same network as SCL:
   #"TIMER".TIMER_1.TON(IN := "AUTOMAT" AND (#STEP_43 = #SQCR), PT := t#500ms);
   IF #"TIMER".TIMER_1.Q THEN #SQCR := #STEP_50; END_IF;
END_REGION

REGION Network 18: STEP 50 ROZHODOVANI Z RECEPTURY CO POSLAT DAL
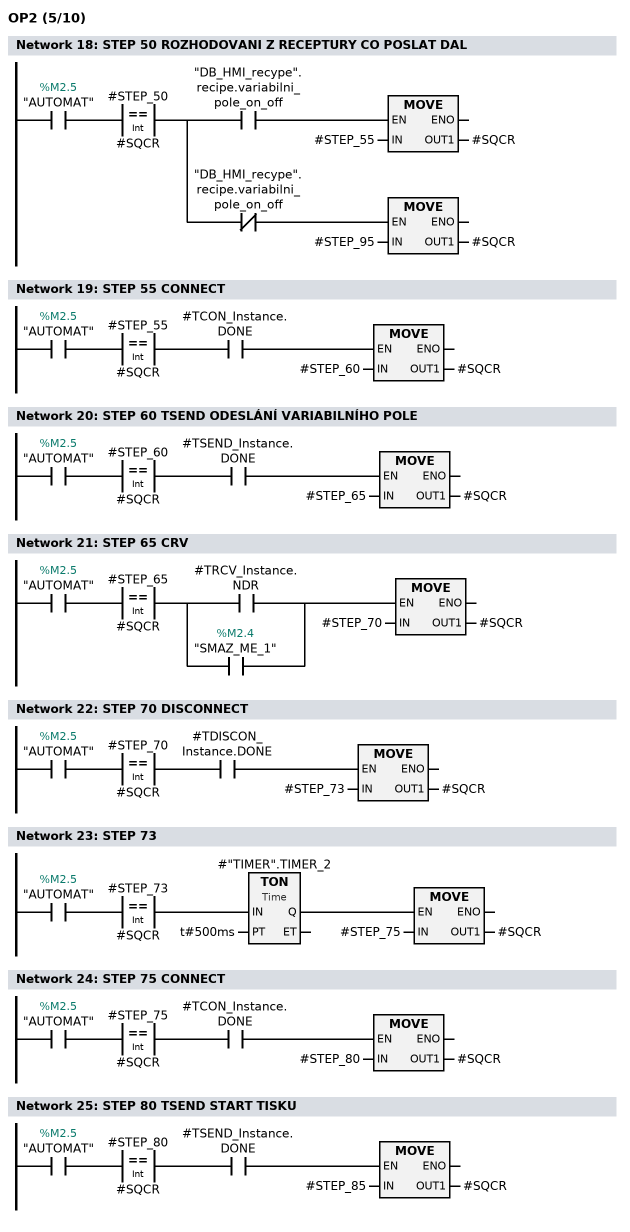
   RUNG wire#powerrail
      Contact( "AUTOMAT" )
      { S7_Templates := "SrcType := Int" } EQ_Contact(in1 := #STEP_50, in2 := #SQCR)
      wire#w1
      Contact( "DB_HMI_recype".recipe.variabilni_pole_on_off )
      Move(in := #STEP_55, out1 => #SQCR)
   END_RUNG
   RUNG wire#w1
      I_Contact( "DB_HMI_recype".recipe.variabilni_pole_on_off )
      Move(in := #STEP_95, out1 => #SQCR)
   END_RUNG
   // the same network as SCL:
   #_w1 := "AUTOMAT" AND (#STEP_50 = #SQCR);
   IF #_w1 AND "DB_HMI_recype".recipe.variabilni_pole_on_off THEN #SQCR := #STEP_55; END_IF;
   IF #_w1 AND NOT "DB_HMI_recype".recipe.variabilni_pole_on_off THEN #SQCR := #STEP_95; END_IF;
END_REGION

REGION Network 19: STEP 55 CONNECT
   RUNG wire#powerrail
      Contact( "AUTOMAT" )
      { S7_Templates := "SrcType := Int" } EQ_Contact(in1 := #STEP_55, in2 := #SQCR)
      Contact( #TCON_Instance.DONE )
      Move(in := #STEP_60, out1 => #SQCR)
   END_RUNG
   // the same network as SCL:
   IF "AUTOMAT" AND (#STEP_55 = #SQCR) AND #TCON_Instance.DONE THEN #SQCR := #STEP_60; END_IF;
END_REGION

REGION Network 20: STEP 60 TSEND ODESLÁNÍ VARIABILNÍHO POLE
   RUNG wire#powerrail
      Contact( "AUTOMAT" )
      { S7_Templates := "SrcType := Int" } EQ_Contact(in1 := #STEP_60, in2 := #SQCR)
      Contact( #TSEND_Instance.DONE )
      Move(in := #STEP_65, out1 => #SQCR)
   END_RUNG
   // the same network as SCL:
   IF "AUTOMAT" AND (#STEP_60 = #SQCR) AND #TSEND_Instance.DONE THEN #SQCR := #STEP_65; END_IF;
END_REGION

REGION Network 21: STEP 65 CRV
   RUNG wire#powerrail
      Contact( "AUTOMAT" )
      { S7_Templates := "SrcType := Int" } EQ_Contact(in1 := #STEP_65, in2 := #SQCR)
      wire#w1
      Contact( #TRCV_Instance.NDR )
      wire#w2
      Move(in := #STEP_70, out1 => #SQCR)
   END_RUNG
   RUNG wire#w1
      Contact( "SMAZ_ME_1" )
   END_RUNG wire#w2
   // the same network as SCL:
   IF "AUTOMAT" AND (#STEP_65 = #SQCR) AND (#TRCV_Instance.NDR OR "SMAZ_ME_1") THEN
       #SQCR := #STEP_70;
   END_IF;
END_REGION

REGION Network 22: STEP 70 DISCONNECT
   RUNG wire#powerrail
      Contact( "AUTOMAT" )
      { S7_Templates := "SrcType := Int" } EQ_Contact(in1 := #STEP_70, in2 := #SQCR)
      Contact( #TDISCON_Instance.DONE )
      Move(in := #STEP_73, out1 => #SQCR)
   END_RUNG
   // the same network as SCL:
   IF "AUTOMAT" AND (#STEP_70 = #SQCR) AND #TDISCON_Instance.DONE THEN #SQCR := #STEP_73; END_IF;
END_REGION

REGION Network 23: STEP 73
   RUNG wire#powerrail
      Contact( "AUTOMAT" )
      { S7_Templates := "SrcType := Int" } EQ_Contact(in1 := #STEP_73, in2 := #SQCR)
      { S7_Templates := "time_type := Time" } #"TIMER".TIMER_2.TON(pt := t#500ms, et =>)
      Move(in := #STEP_75, out1 => #SQCR)
   END_RUNG
   // the same network as SCL:
   #"TIMER".TIMER_2.TON(IN := "AUTOMAT" AND (#STEP_73 = #SQCR), PT := t#500ms);
   IF #"TIMER".TIMER_2.Q THEN #SQCR := #STEP_75; END_IF;
END_REGION

REGION Network 24: STEP 75 CONNECT
   RUNG wire#powerrail
      Contact( "AUTOMAT" )
      { S7_Templates := "SrcType := Int" } EQ_Contact(in1 := #STEP_75, in2 := #SQCR)
      Contact( #TCON_Instance.DONE )
      Move(in := #STEP_80, out1 => #SQCR)
   END_RUNG
   // the same network as SCL:
   IF "AUTOMAT" AND (#STEP_75 = #SQCR) AND #TCON_Instance.DONE THEN #SQCR := #STEP_80; END_IF;
END_REGION

REGION Network 25: STEP 80 TSEND START TISKU
   RUNG wire#powerrail
      Contact( "AUTOMAT" )
      { S7_Templates := "SrcType := Int" } EQ_Contact(in1 := #STEP_80, in2 := #SQCR)
      Contact( #TSEND_Instance.DONE )
      Move(in := #STEP_85, out1 => #SQCR)
   END_RUNG
   // the same network as SCL:
   IF "AUTOMAT" AND (#STEP_80 = #SQCR) AND #TSEND_Instance.DONE THEN #SQCR := #STEP_85; END_IF;
END_REGION

REGION Network 26: STEP 85 TRCV
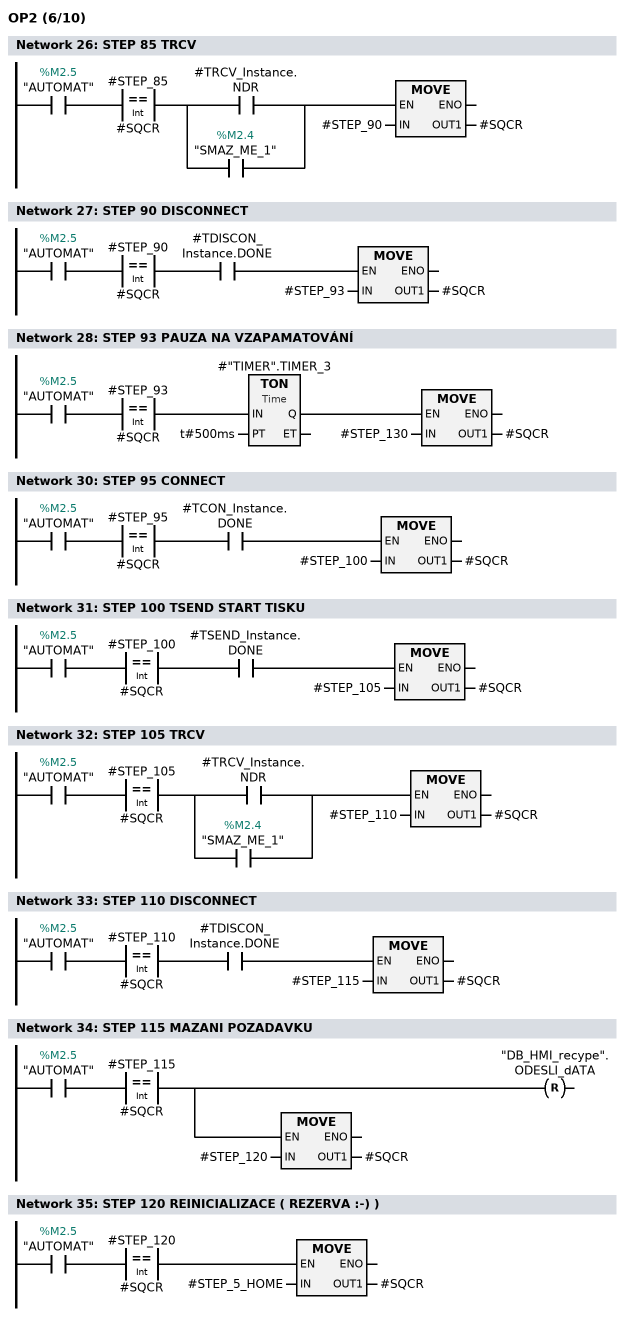
   RUNG wire#powerrail
      Contact( "AUTOMAT" )
      { S7_Templates := "SrcType := Int" } EQ_Contact(in1 := #STEP_85, in2 := #SQCR)
      wire#w1
      Contact( #TRCV_Instance.NDR )
      wire#w2
      Move(in := #STEP_90, out1 => #SQCR)
   END_RUNG
   RUNG wire#w1
      Contact( "SMAZ_ME_1" )
   END_RUNG wire#w2
   // the same network as SCL:
   IF "AUTOMAT" AND (#STEP_85 = #SQCR) AND (#TRCV_Instance.NDR OR "SMAZ_ME_1") THEN
       #SQCR := #STEP_90;
   END_IF;
END_REGION

REGION Network 27: STEP 90 DISCONNECT
   RUNG wire#powerrail
      Contact( "AUTOMAT" )
      { S7_Templates := "SrcType := Int" } EQ_Contact(in1 := #STEP_90, in2 := #SQCR)
      Contact( #TDISCON_Instance.DONE )
      Move(in := #STEP_93, out1 => #SQCR)
   END_RUNG
   // the same network as SCL:
   IF "AUTOMAT" AND (#STEP_90 = #SQCR) AND #TDISCON_Instance.DONE THEN #SQCR := #STEP_93; END_IF;
END_REGION

REGION Network 28: STEP 93 PAUZA NA VZAPAMATOVÁNÍ
   RUNG wire#powerrail
      Contact( "AUTOMAT" )
      { S7_Templates := "SrcType := Int" } EQ_Contact(in1 := #STEP_93, in2 := #SQCR)
      { S7_Templates := "time_type := Time" } #"TIMER".TIMER_3.TON(pt := t#500ms, et =>)
      Move(in := #STEP_130, out1 => #SQCR)
   END_RUNG
   // the same network as SCL:
   #"TIMER".TIMER_3.TON(IN := "AUTOMAT" AND (#STEP_93 = #SQCR), PT := t#500ms);
   IF #"TIMER".TIMER_3.Q THEN #SQCR := #STEP_130; END_IF;
END_REGION

REGION Network 29 (SCL): JEDEN RAMEC
   IF #Tisk.jeden_ramec AND #SQCR = #STEP_130 THEN
       #SQCR := #STEP_95;
   END_IF;
END_REGION

REGION Network 30: STEP 95 CONNECT
   RUNG wire#powerrail
      Contact( "AUTOMAT" )
      { S7_Templates := "SrcType := Int" } EQ_Contact(in1 := #STEP_95, in2 := #SQCR)
      Contact( #TCON_Instance.DONE )
      Move(in := #STEP_100, out1 => #SQCR)
   END_RUNG
   // the same network as SCL:
   IF "AUTOMAT" AND (#STEP_95 = #SQCR) AND #TCON_Instance.DONE THEN #SQCR := #STEP_100; END_IF;
END_REGION

REGION Network 31: STEP 100 TSEND START TISKU
   RUNG wire#powerrail
      Contact( "AUTOMAT" )
      { S7_Templates := "SrcType := Int" } EQ_Contact(in1 := #STEP_100, in2 := #SQCR)
      Contact( #TSEND_Instance.DONE )
      Move(in := #STEP_105, out1 => #SQCR)
   END_RUNG
   // the same network as SCL:
   IF "AUTOMAT" AND (#STEP_100 = #SQCR) AND #TSEND_Instance.DONE THEN #SQCR := #STEP_105; END_IF;
END_REGION

REGION Network 32: STEP 105 TRCV
   RUNG wire#powerrail
      Contact( "AUTOMAT" )
      { S7_Templates := "SrcType := Int" } EQ_Contact(in1 := #STEP_105, in2 := #SQCR)
      wire#w1
      Contact( #TRCV_Instance.NDR )
      wire#w2
      Move(in := #STEP_110, out1 => #SQCR)
   END_RUNG
   RUNG wire#w1
      Contact( "SMAZ_ME_1" )
   END_RUNG wire#w2
   // the same network as SCL:
   IF "AUTOMAT" AND (#STEP_105 = #SQCR) AND (#TRCV_Instance.NDR OR "SMAZ_ME_1") THEN
       #SQCR := #STEP_110;
   END_IF;
END_REGION

REGION Network 33: STEP 110 DISCONNECT
   RUNG wire#powerrail
      Contact( "AUTOMAT" )
      { S7_Templates := "SrcType := Int" } EQ_Contact(in1 := #STEP_110, in2 := #SQCR)
      Contact( #TDISCON_Instance.DONE )
      Move(in := #STEP_115, out1 => #SQCR)
   END_RUNG
   // the same network as SCL:
   IF "AUTOMAT" AND (#STEP_110 = #SQCR) AND #TDISCON_Instance.DONE THEN #SQCR := #STEP_115; END_IF;
END_REGION

REGION Network 34: STEP 115 MAZANI POZADAVKU
   RUNG wire#powerrail
      Contact( "AUTOMAT" )
      { S7_Templates := "SrcType := Int" } EQ_Contact(in1 := #STEP_115, in2 := #SQCR)
      wire#w1
      R_Coil( "DB_HMI_recype".ODESLI_dATA )
   END_RUNG
   RUNG wire#w1
      Move(in := #STEP_120, out1 => #SQCR)
   END_RUNG
   // the same network as SCL:
   IF "AUTOMAT" AND (#STEP_115 = #SQCR) THEN
       "DB_HMI_recype".ODESLI_dATA := FALSE;
       #SQCR := #STEP_120;
   END_IF;
END_REGION

REGION Network 35: STEP 120 REINICIALIZACE ( REZERVA :-) )
   RUNG wire#powerrail
      Contact( "AUTOMAT" )
      { S7_Templates := "SrcType := Int" } EQ_Contact(in1 := #STEP_120, in2 := #SQCR)
      Move(in := #STEP_5_HOME, out1 => #SQCR)
   END_RUNG
   // the same network as SCL:
   IF "AUTOMAT" AND (#STEP_120 = #SQCR) THEN #SQCR := #STEP_5_HOME; END_IF;
END_REGION

REGION Network 36: STEP 130 CONNECT
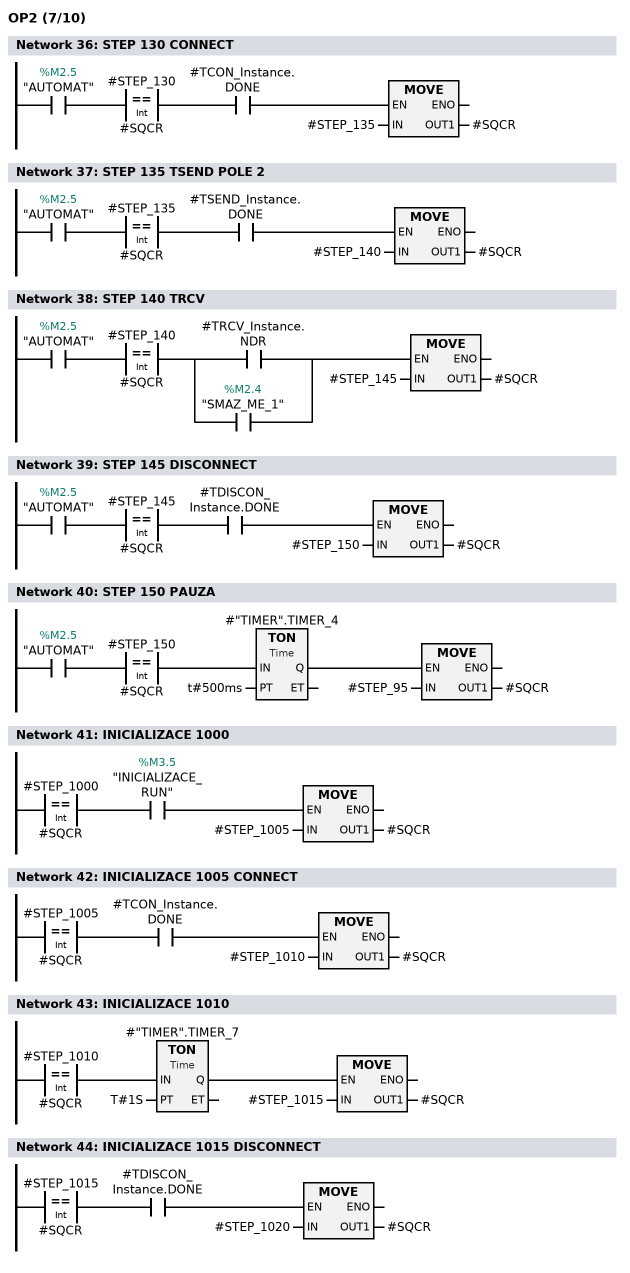
   RUNG wire#powerrail
      Contact( "AUTOMAT" )
      { S7_Templates := "SrcType := Int" } EQ_Contact(in1 := #STEP_130, in2 := #SQCR)
      Contact( #TCON_Instance.DONE )
      Move(in := #STEP_135, out1 => #SQCR)
   END_RUNG
   // the same network as SCL:
   IF "AUTOMAT" AND (#STEP_130 = #SQCR) AND #TCON_Instance.DONE THEN #SQCR := #STEP_135; END_IF;
END_REGION

REGION Network 37: STEP 135 TSEND POLE 2
   RUNG wire#powerrail
      Contact( "AUTOMAT" )
      { S7_Templates := "SrcType := Int" } EQ_Contact(in1 := #STEP_135, in2 := #SQCR)
      Contact( #TSEND_Instance.DONE )
      Move(in := #STEP_140, out1 => #SQCR)
   END_RUNG
   // the same network as SCL:
   IF "AUTOMAT" AND (#STEP_135 = #SQCR) AND #TSEND_Instance.DONE THEN #SQCR := #STEP_140; END_IF;
END_REGION

REGION Network 38: STEP 140 TRCV
   RUNG wire#powerrail
      Contact( "AUTOMAT" )
      { S7_Templates := "SrcType := Int" } EQ_Contact(in1 := #STEP_140, in2 := #SQCR)
      wire#w1
      Contact( #TRCV_Instance.NDR )
      wire#w2
      Move(in := #STEP_145, out1 => #SQCR)
   END_RUNG
   RUNG wire#w1
      Contact( "SMAZ_ME_1" )
   END_RUNG wire#w2
   // the same network as SCL:
   IF "AUTOMAT" AND (#STEP_140 = #SQCR) AND (#TRCV_Instance.NDR OR "SMAZ_ME_1") THEN
       #SQCR := #STEP_145;
   END_IF;
END_REGION

REGION Network 39: STEP 145 DISCONNECT
   RUNG wire#powerrail
      Contact( "AUTOMAT" )
      { S7_Templates := "SrcType := Int" } EQ_Contact(in1 := #STEP_145, in2 := #SQCR)
      Contact( #TDISCON_Instance.DONE )
      Move(in := #STEP_150, out1 => #SQCR)
   END_RUNG
   // the same network as SCL:
   IF "AUTOMAT" AND (#STEP_145 = #SQCR) AND #TDISCON_Instance.DONE THEN #SQCR := #STEP_150; END_IF;
END_REGION

REGION Network 40: STEP 150 PAUZA
   RUNG wire#powerrail
      Contact( "AUTOMAT" )
      { S7_Templates := "SrcType := Int" } EQ_Contact(in1 := #STEP_150, in2 := #SQCR)
      { S7_Templates := "time_type := Time" } #"TIMER".TIMER_4.TON(pt := t#500ms, et =>)
      Move(in := #STEP_95, out1 => #SQCR)
   END_RUNG
   // the same network as SCL:
   #"TIMER".TIMER_4.TON(IN := "AUTOMAT" AND (#STEP_150 = #SQCR), PT := t#500ms);
   IF #"TIMER".TIMER_4.Q THEN #SQCR := #STEP_95; END_IF;
END_REGION

REGION Network 41: INICIALIZACE 1000
   RUNG wire#powerrail
      { S7_Templates := "SrcType := Int" } EQ_Contact(in1 := #STEP_1000, in2 := #SQCR)
      Contact( "INICIALIZACE_RUN" )
      Move(in := #STEP_1005, out1 => #SQCR)
   END_RUNG
   // the same network as SCL:
   IF (#STEP_1000 = #SQCR) AND "INICIALIZACE_RUN" THEN #SQCR := #STEP_1005; END_IF;
END_REGION

REGION Network 42: INICIALIZACE 1005 CONNECT
   RUNG wire#powerrail
      { S7_Templates := "SrcType := Int" } EQ_Contact(in1 := #STEP_1005, in2 := #SQCR)
      Contact( #TCON_Instance.DONE )
      Move(in := #STEP_1010, out1 => #SQCR)
   END_RUNG
   // the same network as SCL:
   IF (#STEP_1005 = #SQCR) AND #TCON_Instance.DONE THEN #SQCR := #STEP_1010; END_IF;
END_REGION

REGION Network 43: INICIALIZACE 1010
   RUNG wire#powerrail
      { S7_Templates := "SrcType := Int" } EQ_Contact(in1 := #STEP_1010, in2 := #SQCR)
      { S7_Templates := "time_type := Time" } #"TIMER".TIMER_7.TON(pt := T#1S, et =>)
      Move(in := #STEP_1015, out1 => #SQCR)
   END_RUNG
   // the same network as SCL:
   #"TIMER".TIMER_7.TON(IN := #STEP_1010 = #SQCR, PT := T#1S);
   IF #"TIMER".TIMER_7.Q THEN #SQCR := #STEP_1015; END_IF;
END_REGION

REGION Network 44: INICIALIZACE 1015 DISCONNECT
   RUNG wire#powerrail
      { S7_Templates := "SrcType := Int" } EQ_Contact(in1 := #STEP_1015, in2 := #SQCR)
      Contact( #TDISCON_Instance.DONE )
      Move(in := #STEP_1020, out1 => #SQCR)
   END_RUNG
   // the same network as SCL:
   IF (#STEP_1015 = #SQCR) AND #TDISCON_Instance.DONE THEN #SQCR := #STEP_1020; END_IF;
END_REGION

REGION Network 45: INICIALIZACE STEP 1015 REZERVA
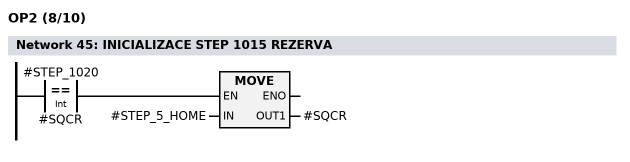
   RUNG wire#powerrail
      { S7_Templates := "SrcType := Int" } EQ_Contact(in1 := #STEP_1020, in2 := #SQCR)
      Move(in := #STEP_5_HOME, out1 => #SQCR)
   END_RUNG
   // the same network as SCL:
   IF #STEP_1020 = #SQCR THEN #SQCR := #STEP_5_HOME; END_IF;
END_REGION

REGION Network 46: automat control door / automat control tiskarna
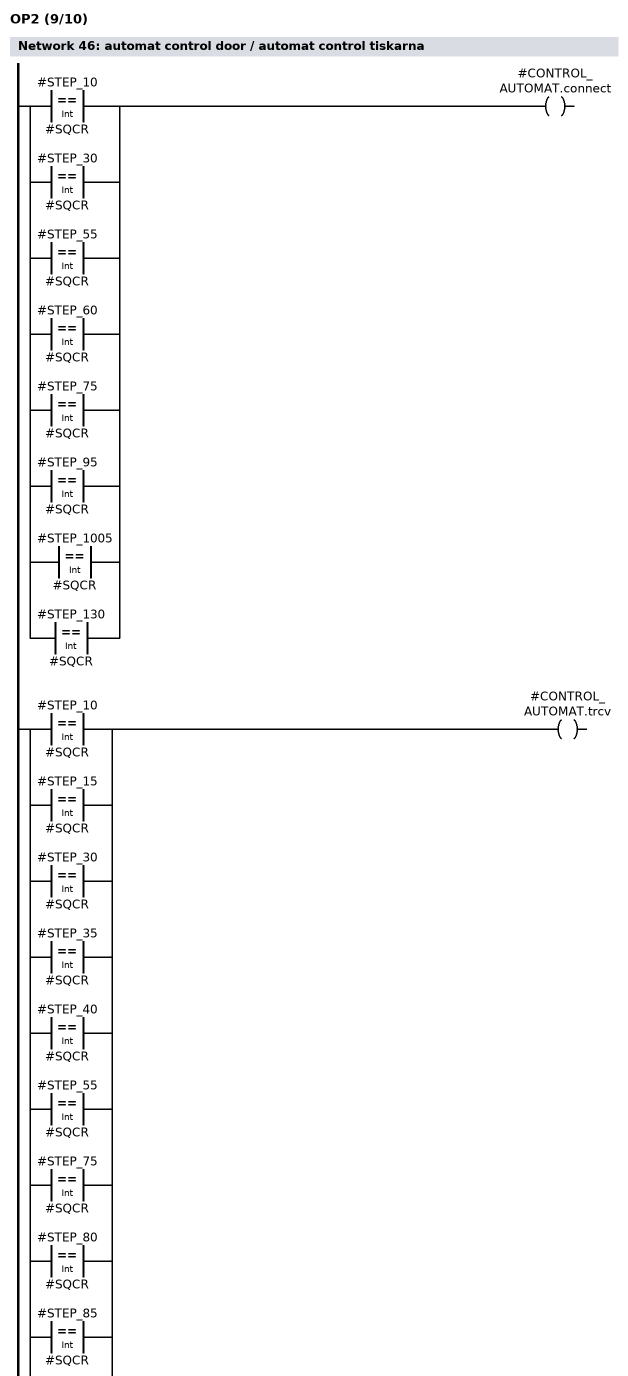
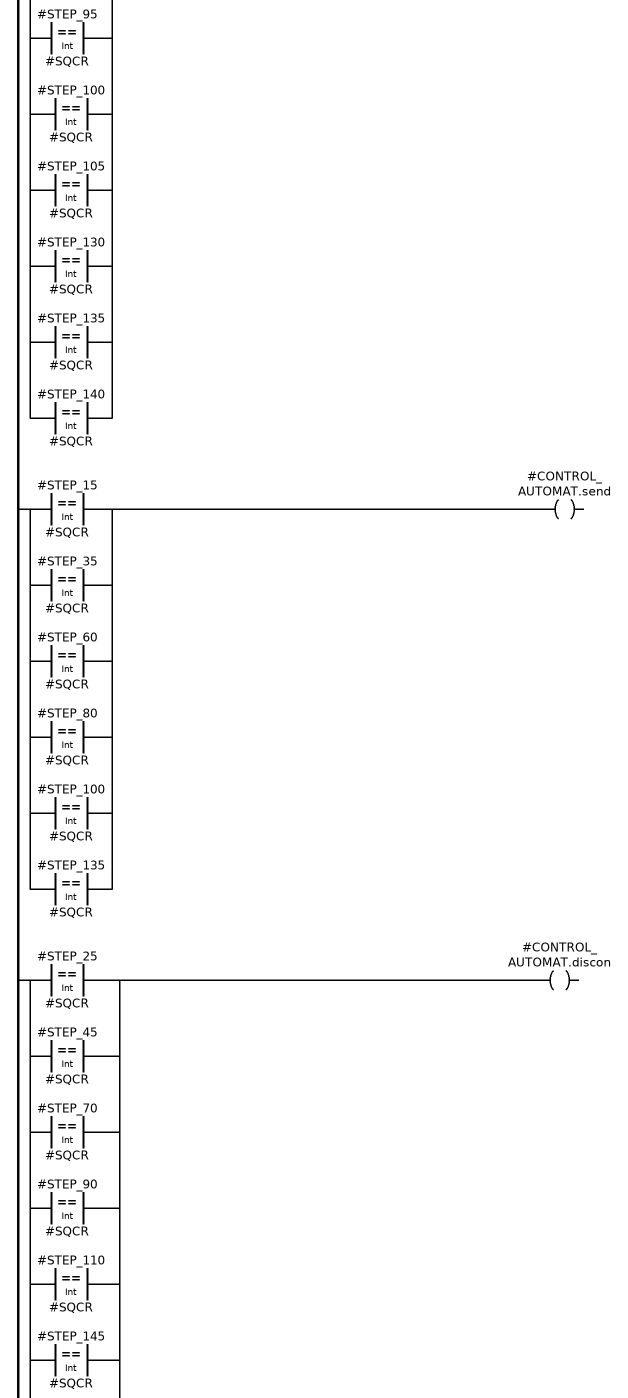
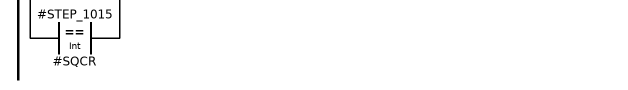
   RUNG wire#powerrail
      { S7_Templates := "SrcType := Int" } EQ_Contact(in1 := #STEP_10, in2 := #SQCR)
      wire#w1
      Coil( #CONTROL_AUTOMAT.connect )
   END_RUNG
   RUNG wire#powerrail
      { S7_Templates := "SrcType := Int" } EQ_Contact(in1 := #STEP_30, in2 := #SQCR)
   END_RUNG wire#w1
   RUNG wire#powerrail
      { S7_Templates := "SrcType := Int" } EQ_Contact(in1 := #STEP_55, in2 := #SQCR)
   END_RUNG wire#w1
   RUNG wire#powerrail
      { S7_Templates := "SrcType := Int" } EQ_Contact(in1 := #STEP_60, in2 := #SQCR)
   END_RUNG wire#w1
   RUNG wire#powerrail
      { S7_Templates := "SrcType := Int" } EQ_Contact(in1 := #STEP_75, in2 := #SQCR)
   END_RUNG wire#w1
   RUNG wire#powerrail
      { S7_Templates := "SrcType := Int" } EQ_Contact(in1 := #STEP_95, in2 := #SQCR)
   END_RUNG wire#w1
   RUNG wire#powerrail
      { S7_Templates := "SrcType := Int" } EQ_Contact(in1 := #STEP_1005, in2 := #SQCR)
   END_RUNG wire#w1
   RUNG wire#powerrail
      { S7_Templates := "SrcType := Int" } EQ_Contact(in1 := #STEP_130, in2 := #SQCR)
   END_RUNG wire#w1
   RUNG wire#powerrail
      { S7_Templates := "SrcType := Int" } EQ_Contact(in1 := #STEP_10, in2 := #SQCR)
      wire#w2
      Coil( #CONTROL_AUTOMAT.trcv )
   END_RUNG
   RUNG wire#powerrail
      { S7_Templates := "SrcType := Int" } EQ_Contact(in1 := #STEP_15, in2 := #SQCR)
   END_RUNG wire#w2
   RUNG wire#powerrail
      { S7_Templates := "SrcType := Int" } EQ_Contact(in1 := #STEP_30, in2 := #SQCR)
   END_RUNG wire#w2
   RUNG wire#powerrail
      { S7_Templates := "SrcType := Int" } EQ_Contact(in1 := #STEP_35, in2 := #SQCR)
   END_RUNG wire#w2
   RUNG wire#powerrail
      { S7_Templates := "SrcType := Int" } EQ_Contact(in1 := #STEP_40, in2 := #SQCR)
   END_RUNG wire#w2
   RUNG wire#powerrail
      { S7_Templates := "SrcType := Int" } EQ_Contact(in1 := #STEP_55, in2 := #SQCR)
   END_RUNG wire#w2
   RUNG wire#powerrail
      { S7_Templates := "SrcType := Int" } EQ_Contact(in1 := #STEP_75, in2 := #SQCR)
   END_RUNG wire#w2
   RUNG wire#powerrail
      { S7_Templates := "SrcType := Int" } EQ_Contact(in1 := #STEP_80, in2 := #SQCR)
   END_RUNG wire#w2
   RUNG wire#powerrail
      { S7_Templates := "SrcType := Int" } EQ_Contact(in1 := #STEP_85, in2 := #SQCR)
   END_RUNG wire#w2
   RUNG wire#powerrail
      { S7_Templates := "SrcType := Int" } EQ_Contact(in1 := #STEP_95, in2 := #SQCR)
   END_RUNG wire#w2
   RUNG wire#powerrail
      { S7_Templates := "SrcType := Int" } EQ_Contact(in1 := #STEP_100, in2 := #SQCR)
   END_RUNG wire#w2
   RUNG wire#powerrail
      { S7_Templates := "SrcType := Int" } EQ_Contact(in1 := #STEP_105, in2 := #SQCR)
   END_RUNG wire#w2
   RUNG wire#powerrail
      { S7_Templates := "SrcType := Int" } EQ_Contact(in1 := #STEP_130, in2 := #SQCR)
   END_RUNG wire#w2
   RUNG wire#powerrail
      { S7_Templates := "SrcType := Int" } EQ_Contact(in1 := #STEP_135, in2 := #SQCR)
   END_RUNG wire#w2
   RUNG wire#powerrail
      { S7_Templates := "SrcType := Int" } EQ_Contact(in1 := #STEP_140, in2 := #SQCR)
   END_RUNG wire#w2
   RUNG wire#powerrail
      { S7_Templates := "SrcType := Int" } EQ_Contact(in1 := #STEP_15, in2 := #SQCR)
      wire#w3
      Coil( #CONTROL_AUTOMAT.send )
   END_RUNG
   RUNG wire#powerrail
      { S7_Templates := "SrcType := Int" } EQ_Contact(in1 := #STEP_35, in2 := #SQCR)
   END_RUNG wire#w3
   RUNG wire#powerrail
      { S7_Templates := "SrcType := Int" } EQ_Contact(in1 := #STEP_60, in2 := #SQCR)
   END_RUNG wire#w3
   RUNG wire#powerrail
      { S7_Templates := "SrcType := Int" } EQ_Contact(in1 := #STEP_80, in2 := #SQCR)
   END_RUNG wire#w3
   RUNG wire#powerrail
      { S7_Templates := "SrcType := Int" } EQ_Contact(in1 := #STEP_100, in2 := #SQCR)
   END_RUNG wire#w3
   RUNG wire#powerrail
      { S7_Templates := "SrcType := Int" } EQ_Contact(in1 := #STEP_135, in2 := #SQCR)
   END_RUNG wire#w3
   RUNG wire#powerrail
      { S7_Templates := "SrcType := Int" } EQ_Contact(in1 := #STEP_25, in2 := #SQCR)
      wire#w4
      Coil( #CONTROL_AUTOMAT.discon )
   END_RUNG
   RUNG wire#powerrail
      { S7_Templates := "SrcType := Int" } EQ_Contact(in1 := #STEP_45, in2 := #SQCR)
   END_RUNG wire#w4
   RUNG wire#powerrail
      { S7_Templates := "SrcType := Int" } EQ_Contact(in1 := #STEP_70, in2 := #SQCR)
   END_RUNG wire#w4
   RUNG wire#powerrail
      { S7_Templates := "SrcType := Int" } EQ_Contact(in1 := #STEP_90, in2 := #SQCR)
   END_RUNG wire#w4
   RUNG wire#powerrail
      { S7_Templates := "SrcType := Int" } EQ_Contact(in1 := #STEP_110, in2 := #SQCR)
   END_RUNG wire#w4
   RUNG wire#powerrail
      { S7_Templates := "SrcType := Int" } EQ_Contact(in1 := #STEP_145, in2 := #SQCR)
   END_RUNG wire#w4
   RUNG wire#powerrail
      { S7_Templates := "SrcType := Int" } EQ_Contact(in1 := #STEP_1015, in2 := #SQCR)
   END_RUNG wire#w4
   // the same network as SCL:
   #CONTROL_AUTOMAT.connect := (#STEP_10 = #SQCR) OR (#STEP_30 = #SQCR) OR (#STEP_55 = #SQCR) OR (#STEP_60 = #SQCR) OR (#STEP_75 = #SQCR) OR (#STEP_95 = #SQCR) OR (#STEP_1005 = #SQCR) OR (#STEP_130 = #SQCR);
   #CONTROL_AUTOMAT.trcv := (#STEP_10 = #SQCR) OR (#STEP_15 = #SQCR) OR (#STEP_30 = #SQCR) OR (#STEP_35 = #SQCR) OR (#STEP_40 = #SQCR) OR (#STEP_55 = #SQCR) OR (#STEP_75 = #SQCR) OR (#STEP_80 = #SQCR) OR (#STEP_85 = #SQCR) OR (#STEP_95 = #SQCR) OR (#STEP_100 = #SQCR) OR (#STEP_105 = #SQCR) OR (#STEP_130 = #SQCR) OR (#STEP_135 = #SQCR) OR (#STEP_140 = #SQCR);
   #CONTROL_AUTOMAT.send := (#STEP_15 = #SQCR) OR (#STEP_35 = #SQCR) OR (#STEP_60 = #SQCR) OR (#STEP_80 = #SQCR) OR (#STEP_100 = #SQCR) OR (#STEP_135 = #SQCR);
   #CONTROL_AUTOMAT.discon := (#STEP_25 = #SQCR) OR (#STEP_45 = #SQCR) OR (#STEP_70 = #SQCR) OR (#STEP_90 = #SQCR) OR (#STEP_110 = #SQCR) OR (#STEP_145 = #SQCR) OR (#STEP_1015 = #SQCR);
END_REGION

REGION Network 47: EXTERNAL_TRIGER
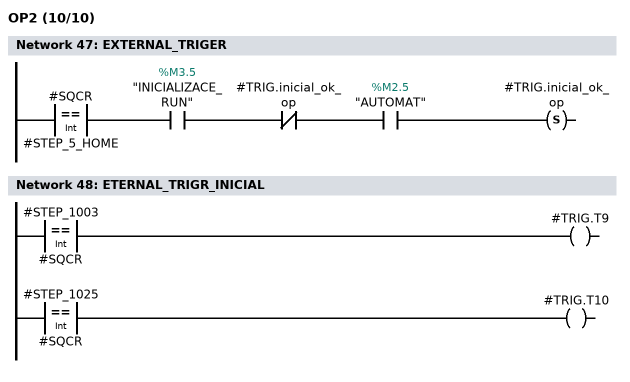
   RUNG wire#powerrail
      { S7_Templates := "SrcType := Int" } EQ_Contact(in1 := #SQCR, in2 := #STEP_5_HOME)
      Contact( "INICIALIZACE_RUN" )
      I_Contact( #TRIG.inicial_ok_op )
      Contact( "AUTOMAT" )
      S_Coil( #TRIG.inicial_ok_op )
   END_RUNG
   // the same network as SCL:
   IF (#SQCR = #STEP_5_HOME) AND "INICIALIZACE_RUN" AND NOT #TRIG.inicial_ok_op AND "AUTOMAT" THEN
       #TRIG.inicial_ok_op := TRUE;
   END_IF;
END_REGION

REGION Network 48: ETERNAL_TRIGR_INICIAL
   RUNG wire#powerrail
      { S7_Templates := "SrcType := Int" } EQ_Contact(in1 := #STEP_1003, in2 := #SQCR)
      Coil( #TRIG.T9 )
   END_RUNG
   RUNG wire#powerrail
      { S7_Templates := "SrcType := Int" } EQ_Contact(in1 := #STEP_1025, in2 := #SQCR)
      Coil( #TRIG.T10 )
   END_RUNG
   // the same network as SCL:
   #TRIG.T9 := #STEP_1003 = #SQCR;
   #TRIG.T10 := #STEP_1025 = #SQCR;
END_REGION

REGION Network 49: hmi
END_REGION
END_FUNCTION_BLOCK

ORGANIZATION_BLOCK "CyclicInterrupt"   // OB30, LAD, CyclicInterrupt
{ S7_Optimized_Access := 'TRUE' }
// stored: SetENOAutomatically false
   VAR_INPUT
      Initial_Call : Bool;   // Initial call of this OB
      Event_Count : Int;   // Events discarded
   END_VAR
   VAR_TEMP
      AKTUALNI_POZICE_FOLIE : DInt;
      AKTUALNI_POZICE_ETIKETA : DInt;
   END_VAR
   VAR_TEMP   // added for the SCL form of the ladder/FBD networks
      _w1 : Bool;
   END_VAR
BEGIN

REGION Network 1
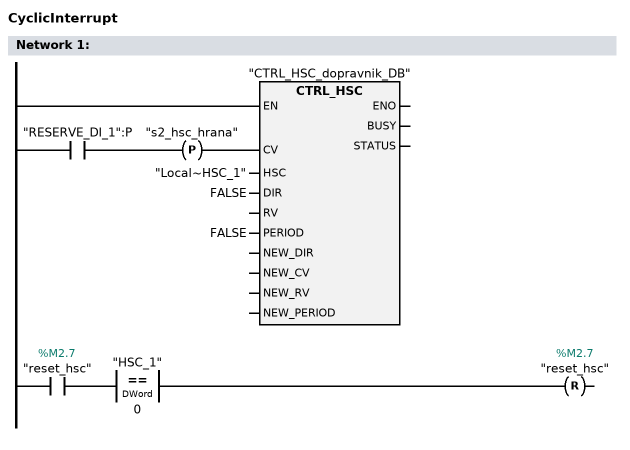
   RUNG wire#powerrail
      "CTRL_HSC_dopravnik_DB".CTRL_HSC(CV := wire#w1, HSC := "Local~HSC_1", DIR := FALSE, RV :=, PERIOD := FALSE, NEW_DIR :=, NEW_CV :=, NEW_RV :=, NEW_PERIOD :=, BUSY =>, STATUS =>)
   END_RUNG
   RUNG wire#powerrail
      Contact( "RESERVE_DI_1":P )
      P_Trig( "s2_hsc_hrana" )
   END_RUNG wire#w1
   RUNG wire#powerrail
      Contact( "reset_hsc" )
      { S7_Templates := "SrcType := DWord" } EQ_Contact(in1 := "HSC_1", in2 := 0)
      R_Coil( "reset_hsc" )
   END_RUNG
   // the same network as SCL:
   #_w1 := "RESERVE_DI_1":P AND NOT "s2_hsc_hrana";   // rising edge
   "s2_hsc_hrana" := "RESERVE_DI_1":P;
   "CTRL_HSC_dopravnik_DB"(CV := #_w1, HSC := "Local~HSC_1", DIR := FALSE, PERIOD := FALSE);   // CTRL_HSC
   IF "reset_hsc" AND ("HSC_1" = 0) THEN "reset_hsc" := FALSE; END_IF;
END_REGION

REGION Network 2 (SCL): Poloha plata od s2 [mm]
   // aktualni_poloha = HSC_1 × mm/puls (fourfold). HSC se nuluje na náběhu s2 (síť 1).
   // Konstanta 1.488 = mm na 1 puls – LIMIT brání přetečení při chodu naprázdno.
   "DB_HMI_recype".aktualni_poloha := REAL_TO_DINT(LIMIT(MN := 0.0,
                                                                                                         IN := DINT_TO_REAL(DWORD_TO_DINT("HSC_1":P)) * 4,
                                                                                                         MX := 99999.0));
END_REGION
END_ORGANIZATION_BLOCK

FUNCTION_BLOCK "OP0"   // FB49, LAD
{ S7_Optimized_Access := 'TRUE' }
// stored: AutoNumber false, MemoryReserve 100, SetENOAutomatically false
   VAR DB_SPECIFIC
      CONTROL_MAN : Struct
         B0 : Bool;
         B1 : Bool;
         B2 : Bool;
         B3 : Bool;
         B4 : Bool;
         B5 : Bool;
         B6 : Bool;
         B7 : Bool;
         B8 : Bool;
         B9 : Bool;
         B10 : Bool;
         B11 : Bool;
         B12 : Bool;
         B13 : Bool;
         B14 : Bool;
         B15 : Bool;
         B16 : Bool;
         B17 : Bool;
         B18 : Bool;
         B19 : Bool;
         B20 : Bool;
         B21 : Bool;
         B22 : Bool;
         B23 : Bool;
         B24 : Bool;
         B25 : Bool;
         B26 : Bool;
         B27 : Bool;
         B28 : Bool;
         B29 : Bool;
         B30 : Bool;
         B31 : Bool;
      END_STRUCT;
      CONTROL_AUTOMAT : Struct
         B0 : Bool;
         B1 : Bool;
         B2 : Bool;
         B3 : Bool;
         B4 : Bool;
         B5 : Bool;
         B6 : Bool;
         B7 : Bool;
         B8 : Bool;
         B9 : Bool;
         B10 : Bool;
         B11 : Bool;
         B12 : Bool;
         B13 : Bool;
         B14 : Bool;
         B15 : Bool;
         B16 : Bool;
         B17 : Bool;
         B18 : Bool;
         B19 : Bool;
         B20 : Bool;
         B21 : Bool;
         B22 : Bool;
         B23 : Bool;
         B24 : Bool;
         B25 : Bool;
         B26 : Bool;
         B27 : Bool;
         B28 : Bool;
         B29 : Bool;
         B30 : Bool;
         B31 : Bool;
      END_STRUCT;
      SENSORS : Struct
         S0 : Bool;
         S1 : Bool;
         S2 : Bool;
         S3 : Bool;
         S4 : Bool;
         S5 : Bool;
         S6 : Bool;
         S7 : Bool;
         S8 : Bool;
         S9 : Bool;
         S10 : Bool;
         S11 : Bool;
         S12 : Bool;
         S13 : Bool;
         S14 : Bool;
         S15 : Bool;
         S16 : Bool;
         S17 : Bool;
         S18 : Bool;
         S19 : Bool;
         S20 : Bool;
         S21 : Bool;
         S22 : Bool;
         S23 : Bool;
         S24 : Bool;
         S25 : Bool;
         S26 : Bool;
         S27 : Bool;
         S28 : Bool;
         S29 : Bool;
         S30 : Bool;
         S31 : Bool;
      END_STRUCT;
      SENSORS_1 : Struct
         S0 : Bool;
         S1 : Bool;
         S2 : Bool;
         S3 : Bool;
         S4 : Bool;
         S5 : Bool;
         S6 : Bool;
         S7 : Bool;
         S8 : Bool;
         S9 : Bool;
         S10 : Bool;
         S11 : Bool;
         S12 : Bool;
         S13 : Bool;
         S14 : Bool;
         S15 : Bool;
         S16 : Bool;
         S17 : Bool;
         S18 : Bool;
         S19 : Bool;
         S20 : Bool;
         S21 : Bool;
         S22 : Bool;
         S23 : Bool;
         S24 : Bool;
         S25 : Bool;
         S26 : Bool;
         S27 : Bool;
         S28 : Bool;
         S29 : Bool;
         S30 : Bool;
         S31 : Bool;
      END_STRUCT;
   END_VAR
   VAR
      S_0 : "SENSOR";
      S_1 { S7_SetPoint := 'True'} : "SENSOR";
      S_2 { S7_SetPoint := 'True'} : "SENSOR";
      S_3 { S7_SetPoint := 'True'} : "SENSOR";
      S_4 { S7_SetPoint := 'True'} : "SENSOR";
      S_5 { S7_SetPoint := 'True'} : "SENSOR";
      S_6 { S7_SetPoint := 'True'} : "SENSOR";
      S_7 { S7_SetPoint := 'True'} : "SENSOR";
      S_8 { S7_SetPoint := 'True'} : "SENSOR";
      S_9 { S7_SetPoint := 'True'} : "SENSOR";
      s_10 { S7_SetPoint := 'True'} : "SENSOR";
      S_11 { S7_SetPoint := 'True'} : "SENSOR";
      S_12 { S7_SetPoint := 'True'} : "SENSOR";
      S_13 { S7_SetPoint := 'True'} : "SENSOR";
      S_14 { S7_SetPoint := 'True'} : "SENSOR";
      S_15 { S7_SetPoint := 'True'} : "SENSOR";
      S_16 { S7_SetPoint := 'True'} : "SENSOR";
      S_17 { S7_SetPoint := 'True'} : "SENSOR";
      S_18 { S7_SetPoint := 'True'} : "SENSOR";
      S_19 { S7_SetPoint := 'True'} : "SENSOR";
      S_20 { S7_SetPoint := 'True'} : "SENSOR";
      S_21 { S7_SetPoint := 'True'} : "SENSOR";
      S_22 { S7_SetPoint := 'True'} : "SENSOR";
      S_23 { S7_SetPoint := 'True'} : "SENSOR";
      S_24 { S7_SetPoint := 'True'} : "SENSOR";
      S_25 { S7_SetPoint := 'True'} : "SENSOR";
      S_26 { S7_SetPoint := 'True'} : "SENSOR";
      S_27 { S7_SetPoint := 'True'} : "SENSOR";
      S_28 { S7_SetPoint := 'True'} : "SENSOR";
      S_29 { S7_SetPoint := 'True'} : "SENSOR";
      S_30 { S7_SetPoint := 'True'} : "SENSOR";
      S_31 { S7_SetPoint := 'True'} : "SENSOR";
      S_32 { S7_SetPoint := 'True'} : "SENSOR";
      S_33 { S7_SetPoint := 'True'} : "SENSOR";
      S_34 { S7_SetPoint := 'True'} : "SENSOR";
      S_35 { S7_SetPoint := 'True'} : "SENSOR";
      M_0 : "MOTOR_CONTROL_BLOCK";
      M_1 { S7_SetPoint := 'True'} : "MOTOR_CONTROL_BLOCK";
      M_2 { S7_SetPoint := 'True'} : "MOTOR_CONTROL_BLOCK";
      M_3 { S7_SetPoint := 'True'} : "MOTOR_CONTROL_BLOCK";
   END_VAR
   VAR DB_SPECIFIC
      SQCR { S7_SetPoint := 'True'} : Int;
      TRIG : Struct
         inicial_ok_op : Bool;
         DSSAD : Bool;
         INICIALIZACE_PROBEHLA : Bool;
         trig_dil : Bool;
         p_trig_control_tcon : Bool;
         T6 : Bool;
         T7 : Bool;
         T8 : Bool;
         T9 : Bool;
         T10 : Bool;
         T11 : Bool;
         T12 : Bool;
         T13 : Bool;
         T14 : Bool;
         T15 : Bool;
         T16 : Bool;
         T17 : Bool;
      END_STRUCT;
      MEMOR : Struct
         M0 : Bool;
         M1 : Bool;
         M2 : Bool;
         M3 : Bool;
         M4 : Bool;
         M5 : Bool;
         M6 : Bool;
         M7 : Bool;
         M8 : Bool;
         M9 : Bool;
         M10 : Bool;
         M11 : Bool;
         RESET_ERROR : Bool;
         M13 : Bool;
         M14 : Bool;
         M15 : Bool;
         M16 : Bool;
         M17 : Bool;
         M18 : Bool;
         M19 : Bool;
         M20 : Bool;
         M21 : Bool;
         M22 : Bool;
         M23 : Bool;
         M24 : Bool;
         M25 : Bool;
         M26 : Bool;
         M27 : Bool;
         M28 : Bool;
         M29 : Bool;
         M30 : Bool;
         M31 : Bool;
         M32 : Bool;
         M33 : Bool;
         start_caklu : Bool;
         M35 : Bool;
         M36 : Bool;
         M37 : Bool;
         M38 : Bool;
         M39 : Bool;
         ALARM_GLOBAL : Bool;
         M41 : Bool;
         M42 : Bool;
         M43 : Bool;
         M44 : Bool;
         M45 : Bool;
         M46 : Bool;
         M47 : Bool;
         M48 : Bool;
         M49 : Bool;
         M50 : Bool;
         M51 : Bool;
         M52 : Bool;
         M53 : Bool;
         M54 : Bool;
         M55 : Bool;
         M56 : Bool;
         M57 : Bool;
         M58 : Bool;
         M59 : Bool;
         M60 : Bool;
         M61 : Bool;
         M62 : Bool;
         M63 : Bool;
      END_STRUCT;
      "TIMER" : Struct
         TIMER_0 : IEC_TIMER;
         TIMER_VACUUM_CLEANER : IEC_TIMER;
         TIMER_DELAY_RESET_EXECUTE : IEC_TIMER;
         TIMER_3 : IEC_TIMER;
         TIMER_4 : IEC_TIMER;
         TIMER_5 : IEC_TIMER;
         TIMER_6 : IEC_TIMER;
         TIMER_7 : IEC_TIMER;
      END_STRUCT;
      HMI : Struct
         povoleni_volby_receptu : Bool;
         "svetlo_on/off" : Bool;
         ALARM_VIDITELNOST : Bool;
         hmi_3 : Bool;
         hmi_4 : Bool;
         hmi_5 : Bool;
         hmi_6 : Bool;
         hmi_7 : Bool;
         hmi_8 : Bool;
         hmi_9 : Bool;
         hmi_10 : Bool;
         hmi_11 : Bool;
         hmi_12 : Bool;
         hmi_13 : Bool;
         hmi_14 : Bool;
         hmi_15 : Bool;
      END_STRUCT;
   END_VAR
   VAR
      kontrola_tcon : Int;
      cyklus_aretace : Int;
      string_pam : String;
      error_m1 : Int;
      error_m2 : Int;
      MAXA : Struct
         ACTUAL_MESSAGE : String[16];
         name_char : Array[0..16] of Char;
         adresace : Byte;
      END_STRUCT;
      HMI_SPEED : Real;
      hmi_man_cab : Bool;
      HMI_START : Bool;
      TRIGR_LASER : DWord;
   END_VAR
   VAR_TEMP
      DATA : Array[0..255] of Char;
      PREVOD : Int;
      NORM_SCALE : LReal;
   END_VAR
   VAR CONSTANT
      STEP_0 : Int := 0;
      step_2 : Int := 2;
      STEP_4 : Int := 4;
      STEP_5_HOME : Int := 5;
      STEP_7 : Int := 7;
      STEP_10 : Int := 10;
      STEP_15 : Int := 15;
      STEP_20 : Int := 20;
      STEP_23 : Int := 23;
      STEP_25 : Int := 25;
      STEP_27 : Int := 27;
      STEP_30 : Int := 30;
      STEP_35 : Int := 35;
      STEP_37 : Int := 37;
      STEP_40 : Int := 40;
      STEP_45 : Int := 45;
      STEP_50 : Int := 50;
      STEP_55 : Int := 55;
      STEP_60 : Int := 60;
      STEP_65 : Int := 65;
      STEP_70 : Int := 70;
      STEP_75 : Int := 75;
      STEP_80 : Int := 80;
      STEP_83 : Int := 83;
      STEP_85 : Int := 85;
      STEP_90 : Int := 90;
      STEP_95 : Int := 95;
      STEP_100 : Int := 100;
      STEP_105 : Int := 105;
      STEP_110 : Int := 110;
      STEP_113 : Int := 113;
      STEP_115 : Int := 115;
      STEP_120 : Int := 120;
      STEP_125 : Int := 125;
      STEP_130 : Int := 130;
      STEP_135 : Int := 135;
      STEP_140 : Int := 140;
      STEP_145 : Int := 145;
      STEP_150 : Int := 150;
      STEP_155 : Int := 155;
      STEP_1000_KONTROLA : Int := 1000;
      STEP_1005_START_INICIAL : Int := 1005;
      STEP_1010_close_door : Int := 1010;
      STEP_1015 : Int := 1015;
      STEP_1020_HOME_OK : Int := 1020;
      STEP_1025 : Int := 1025;
      STEP_3000 : Int := 3000;
      STEP_3005 : Int := 3005;
      STEP_3010 : Int := 3010;
      STEP_3015 : Int := 3015;
      STEP_3020 : Int := 3020;
      STEP_2000 : Int := 2000;
      string_null : String;
      char_null : Char;
   END_VAR
   VAR_TEMP   // added for the SCL form of the ladder/FBD networks
      _w1 : Bool;
      _w2 : Bool;
      _w3 : Bool;
      _w4 : Bool;
      _w5 : Bool;
      _w6 : Bool;
      _w7 : Bool;
      _w8 : Bool;
      _w9 : Bool;
   END_VAR
BEGIN

REGION Network 1 (SCL)
   IF "FirstScan" = true THEN
       #MAXA.adresace := 0;
   END_IF;
     (*  

   #MAXA.name_char[0] := "-XT500_name_byte_0";
   #MAXA.name_char[1] := "-XT500_name_byte_1";
   #MAXA.name_char[2] := "-XT500_name_byte_2";
   #MAXA.name_char[3] := "-XT500_name_byte_3";
   #MAXA.name_char[4] := "-XT500_name_byte_4";
   #MAXA.name_char[5] := "-XT500_name_byte_5";
   #MAXA.name_char[6] := "-XT500_name_byte_6";
   #MAXA.name_char[7] := "-XT500_name_byte_7";
   #MAXA.name_char[8] := "-XT500_name_byte_8";
   #MAXA.name_char[9] := "-XT500_name_byte_9";
   #MAXA.name_char[10] := "-XT500_name_byte_10";
   #MAXA.name_char[11] := "-XT500_name_byte_11";
   #MAXA.name_char[12] := "-XT500_name_byte_12";
   #MAXA.name_char[13] := "-XT500_name_byte_13";
   #MAXA.name_char[14] := "-XT500_name_byte_14";
   #MAXA.name_char[15] := "-XT500_name_byte_15";
   *)

   IF #SQCR <> 0 THEN
       IF #MAXA.adresace > 16 THEN
           #MAXA.adresace := 0;
       END_IF;
       #MAXA.ACTUAL_MESSAGE[#MAXA.adresace + 1] := #MAXA.name_char[#MAXA.adresace];
       #MAXA.adresace := #MAXA.adresace + 1;
   END_IF;
END_REGION

REGION Network 2: manuali ovladani reset
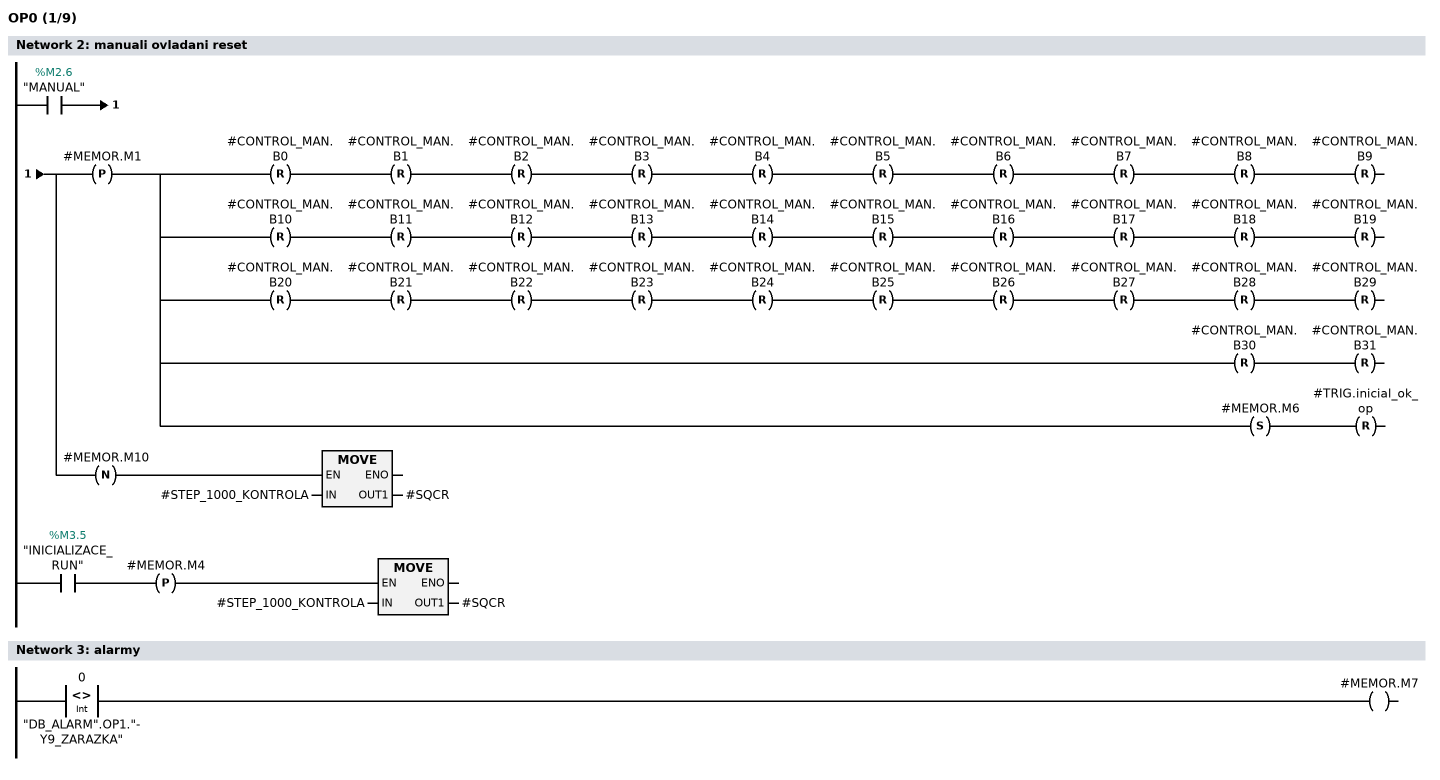
   RUNG wire#powerrail
      Contact( "MANUAL" )
      wire#w1
      P_Trig( #MEMOR.M1 )
      wire#w2
      R_Coil( #CONTROL_MAN.B0 )
      R_Coil( #CONTROL_MAN.B1 )
      R_Coil( #CONTROL_MAN.B2 )
      R_Coil( #CONTROL_MAN.B3 )
      R_Coil( #CONTROL_MAN.B4 )
      R_Coil( #CONTROL_MAN.B5 )
      R_Coil( #CONTROL_MAN.B6 )
      R_Coil( #CONTROL_MAN.B7 )
      R_Coil( #CONTROL_MAN.B8 )
      R_Coil( #CONTROL_MAN.B9 )
   END_RUNG
   RUNG wire#w2
      R_Coil( #CONTROL_MAN.B10 )
      R_Coil( #CONTROL_MAN.B11 )
      R_Coil( #CONTROL_MAN.B12 )
      R_Coil( #CONTROL_MAN.B13 )
      R_Coil( #CONTROL_MAN.B14 )
      R_Coil( #CONTROL_MAN.B15 )
      R_Coil( #CONTROL_MAN.B16 )
      R_Coil( #CONTROL_MAN.B17 )
      R_Coil( #CONTROL_MAN.B18 )
      R_Coil( #CONTROL_MAN.B19 )
   END_RUNG
   RUNG wire#w2
      R_Coil( #CONTROL_MAN.B20 )
      R_Coil( #CONTROL_MAN.B21 )
      R_Coil( #CONTROL_MAN.B22 )
      R_Coil( #CONTROL_MAN.B23 )
      R_Coil( #CONTROL_MAN.B24 )
      R_Coil( #CONTROL_MAN.B25 )
      R_Coil( #CONTROL_MAN.B26 )
      R_Coil( #CONTROL_MAN.B27 )
      R_Coil( #CONTROL_MAN.B28 )
      R_Coil( #CONTROL_MAN.B29 )
   END_RUNG
   RUNG wire#w2
      R_Coil( #CONTROL_MAN.B30 )
      R_Coil( #CONTROL_MAN.B31 )
   END_RUNG
   RUNG wire#w2
      S_Coil( #MEMOR.M6 )
      R_Coil( #TRIG.inicial_ok_op )
   END_RUNG
   RUNG wire#w1
      N_Trig( #MEMOR.M10 )
      Move(in := #STEP_1000_KONTROLA, out1 => #SQCR)
   END_RUNG
   RUNG wire#powerrail
      Contact( "INICIALIZACE_RUN" )
      P_Trig( #MEMOR.M4 )
      Move(in := #STEP_1000_KONTROLA, out1 => #SQCR)
   END_RUNG
   // the same network as SCL:
   #_w1 := "MANUAL" AND NOT #MEMOR.M1;   // rising edge
   #MEMOR.M1 := "MANUAL";
   IF #_w1 THEN
       #CONTROL_MAN.B0 := FALSE;
       #CONTROL_MAN.B1 := FALSE;
       #CONTROL_MAN.B2 := FALSE;
       #CONTROL_MAN.B3 := FALSE;
       #CONTROL_MAN.B4 := FALSE;
       #CONTROL_MAN.B5 := FALSE;
       #CONTROL_MAN.B6 := FALSE;
       #CONTROL_MAN.B7 := FALSE;
       #CONTROL_MAN.B8 := FALSE;
       #CONTROL_MAN.B9 := FALSE;
       #CONTROL_MAN.B10 := FALSE;
       #CONTROL_MAN.B11 := FALSE;
       #CONTROL_MAN.B12 := FALSE;
       #CONTROL_MAN.B13 := FALSE;
       #CONTROL_MAN.B14 := FALSE;
       #CONTROL_MAN.B15 := FALSE;
       #CONTROL_MAN.B16 := FALSE;
       #CONTROL_MAN.B17 := FALSE;
       #CONTROL_MAN.B18 := FALSE;
       #CONTROL_MAN.B19 := FALSE;
       #CONTROL_MAN.B20 := FALSE;
       #CONTROL_MAN.B21 := FALSE;
       #CONTROL_MAN.B22 := FALSE;
       #CONTROL_MAN.B23 := FALSE;
       #CONTROL_MAN.B24 := FALSE;
       #CONTROL_MAN.B25 := FALSE;
       #CONTROL_MAN.B26 := FALSE;
       #CONTROL_MAN.B27 := FALSE;
       #CONTROL_MAN.B28 := FALSE;
       #CONTROL_MAN.B29 := FALSE;
       #CONTROL_MAN.B30 := FALSE;
       #CONTROL_MAN.B31 := FALSE;
       #MEMOR.M6 := TRUE;
       #TRIG.inicial_ok_op := FALSE;
   END_IF;
   #_w2 := NOT "MANUAL" AND #MEMOR.M10;   // falling edge
   #MEMOR.M10 := "MANUAL";
   IF #_w2 THEN #SQCR := #STEP_1000_KONTROLA; END_IF;
   #_w3 := "INICIALIZACE_RUN" AND NOT #MEMOR.M4;   // rising edge
   #MEMOR.M4 := "INICIALIZACE_RUN";
   IF #_w3 THEN #SQCR := #STEP_1000_KONTROLA; END_IF;
END_REGION

REGION Network 3: alarmy
   RUNG wire#powerrail
      { S7_Templates := "SrcType := Int" } NE_Contact(in1 := 0, in2 := "DB_ALARM".OP1."-Y9_ZARAZKA")
      Coil( #MEMOR.M7 )
   END_RUNG
   // the same network as SCL:
   #MEMOR.M7 := 0 <> "DB_ALARM".OP1."-Y9_ZARAZKA";
END_REGION

REGION Network 4: senzory
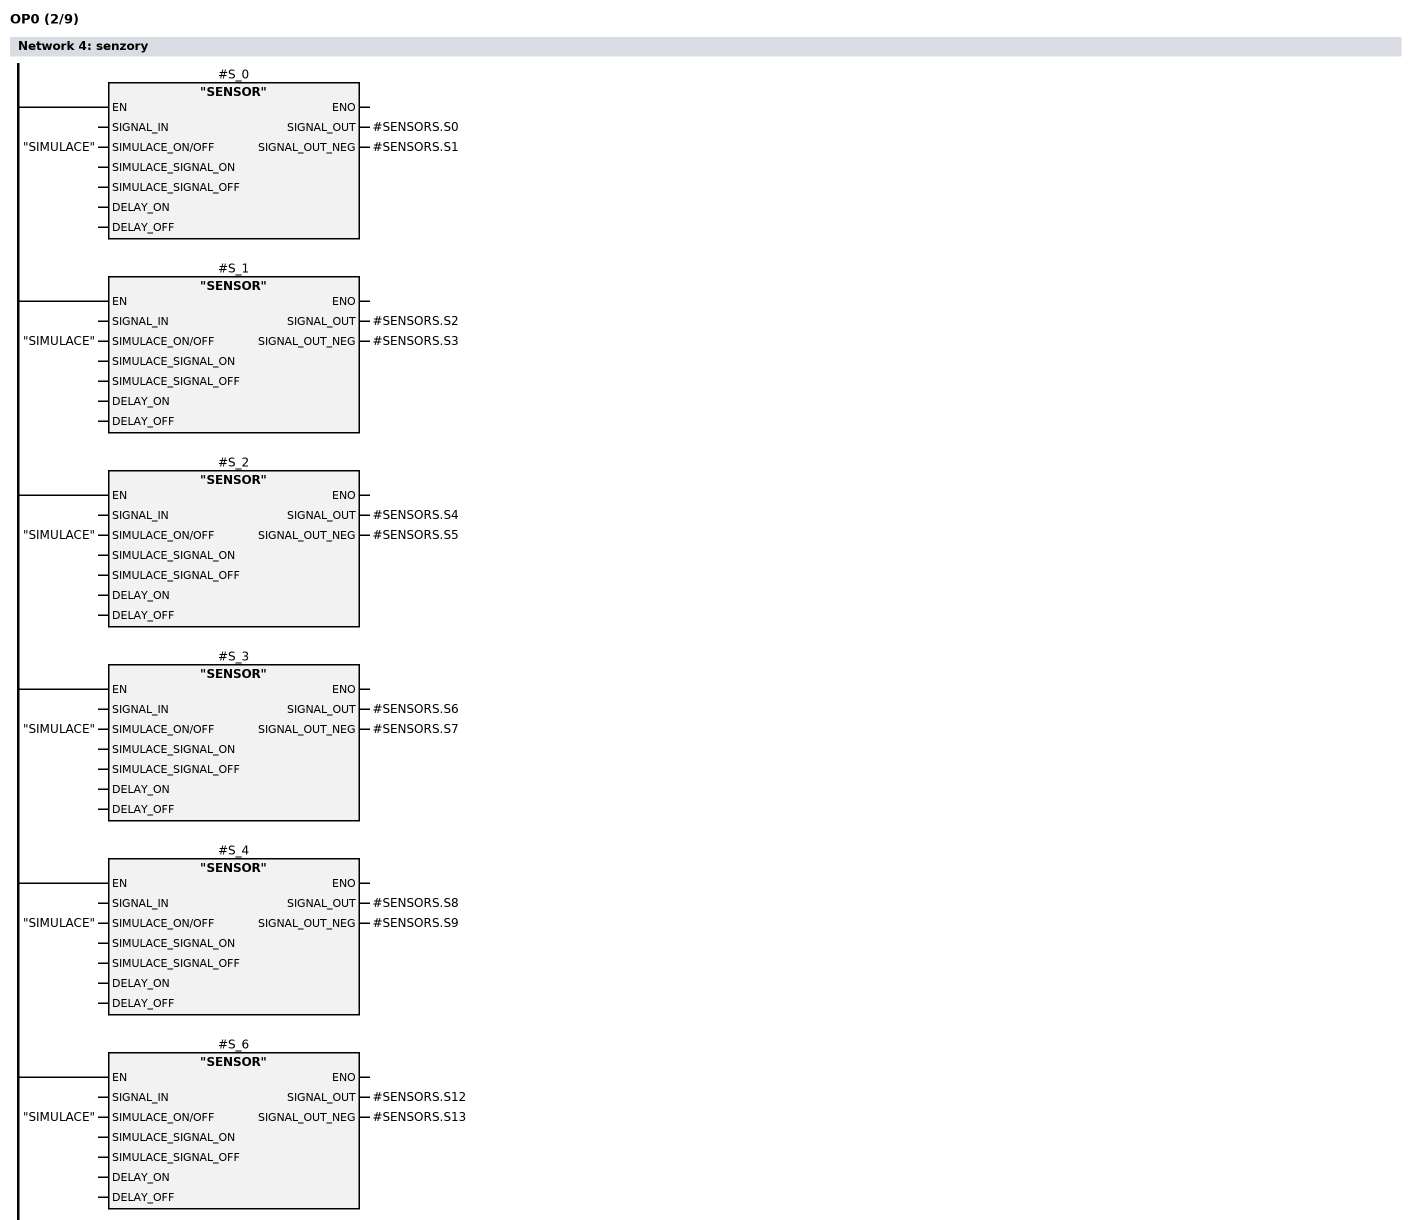
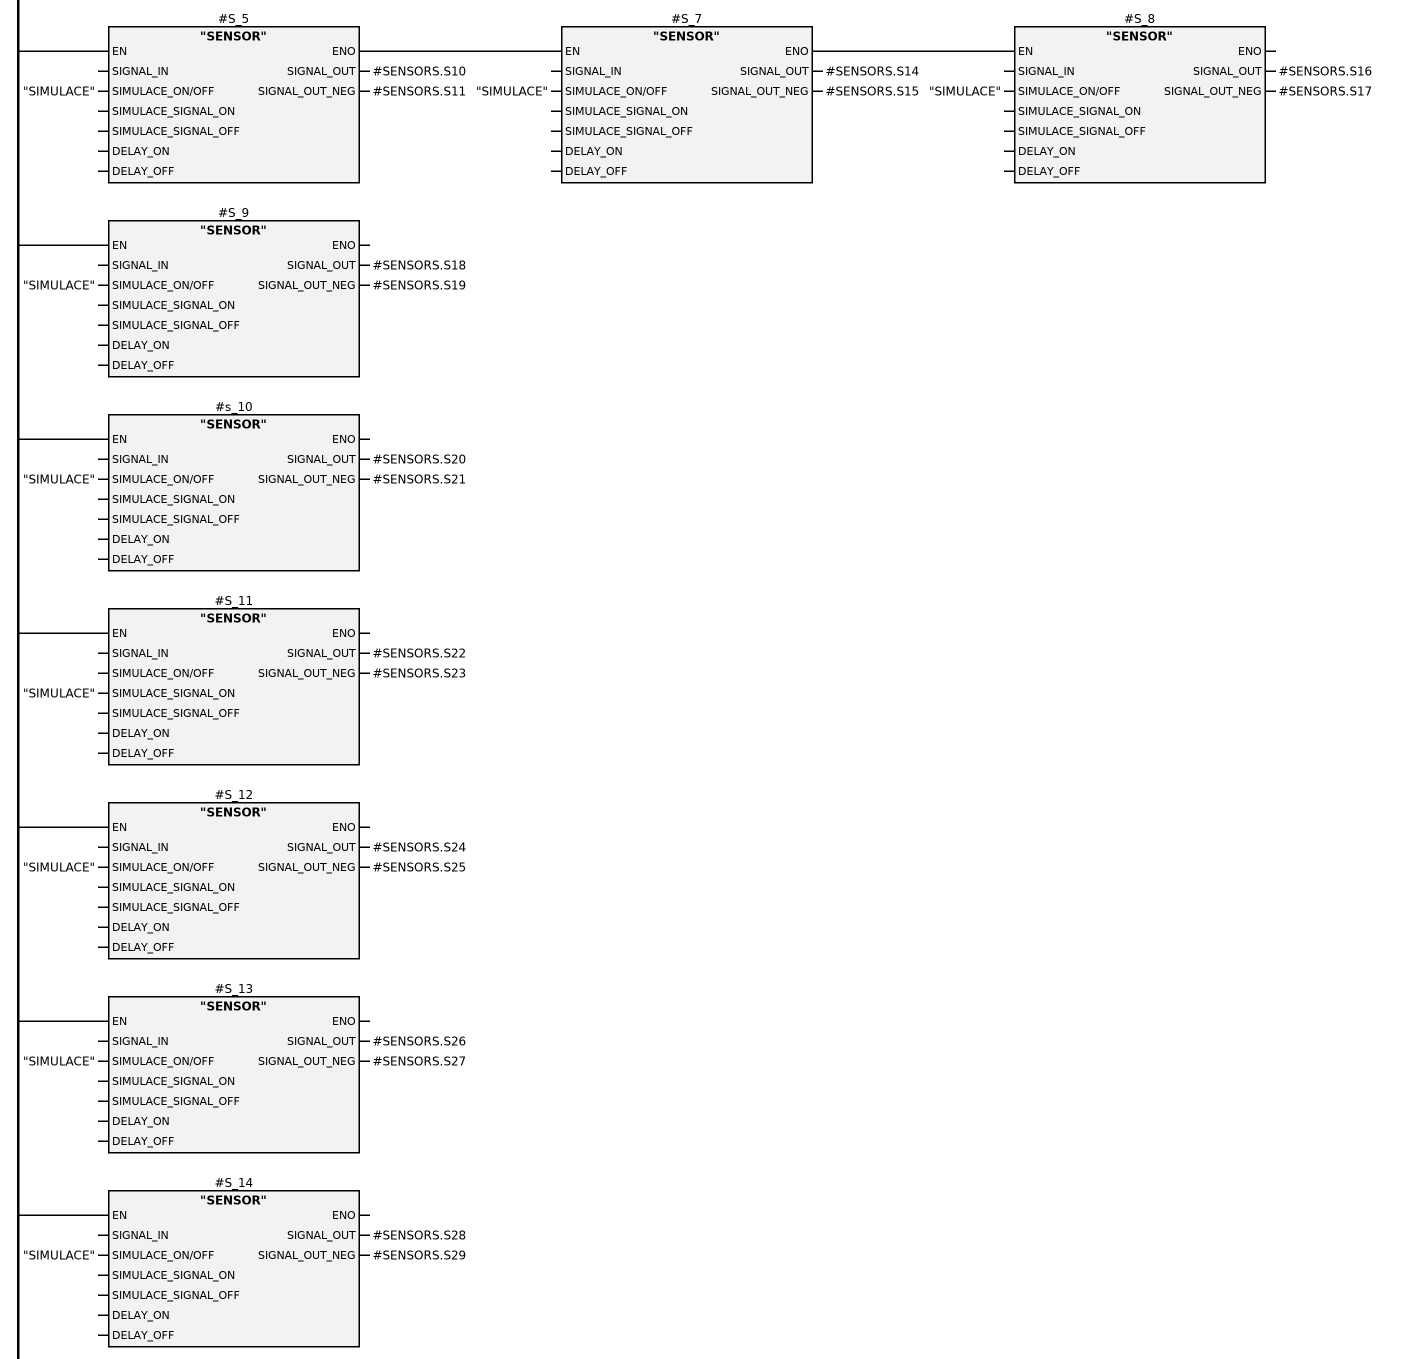
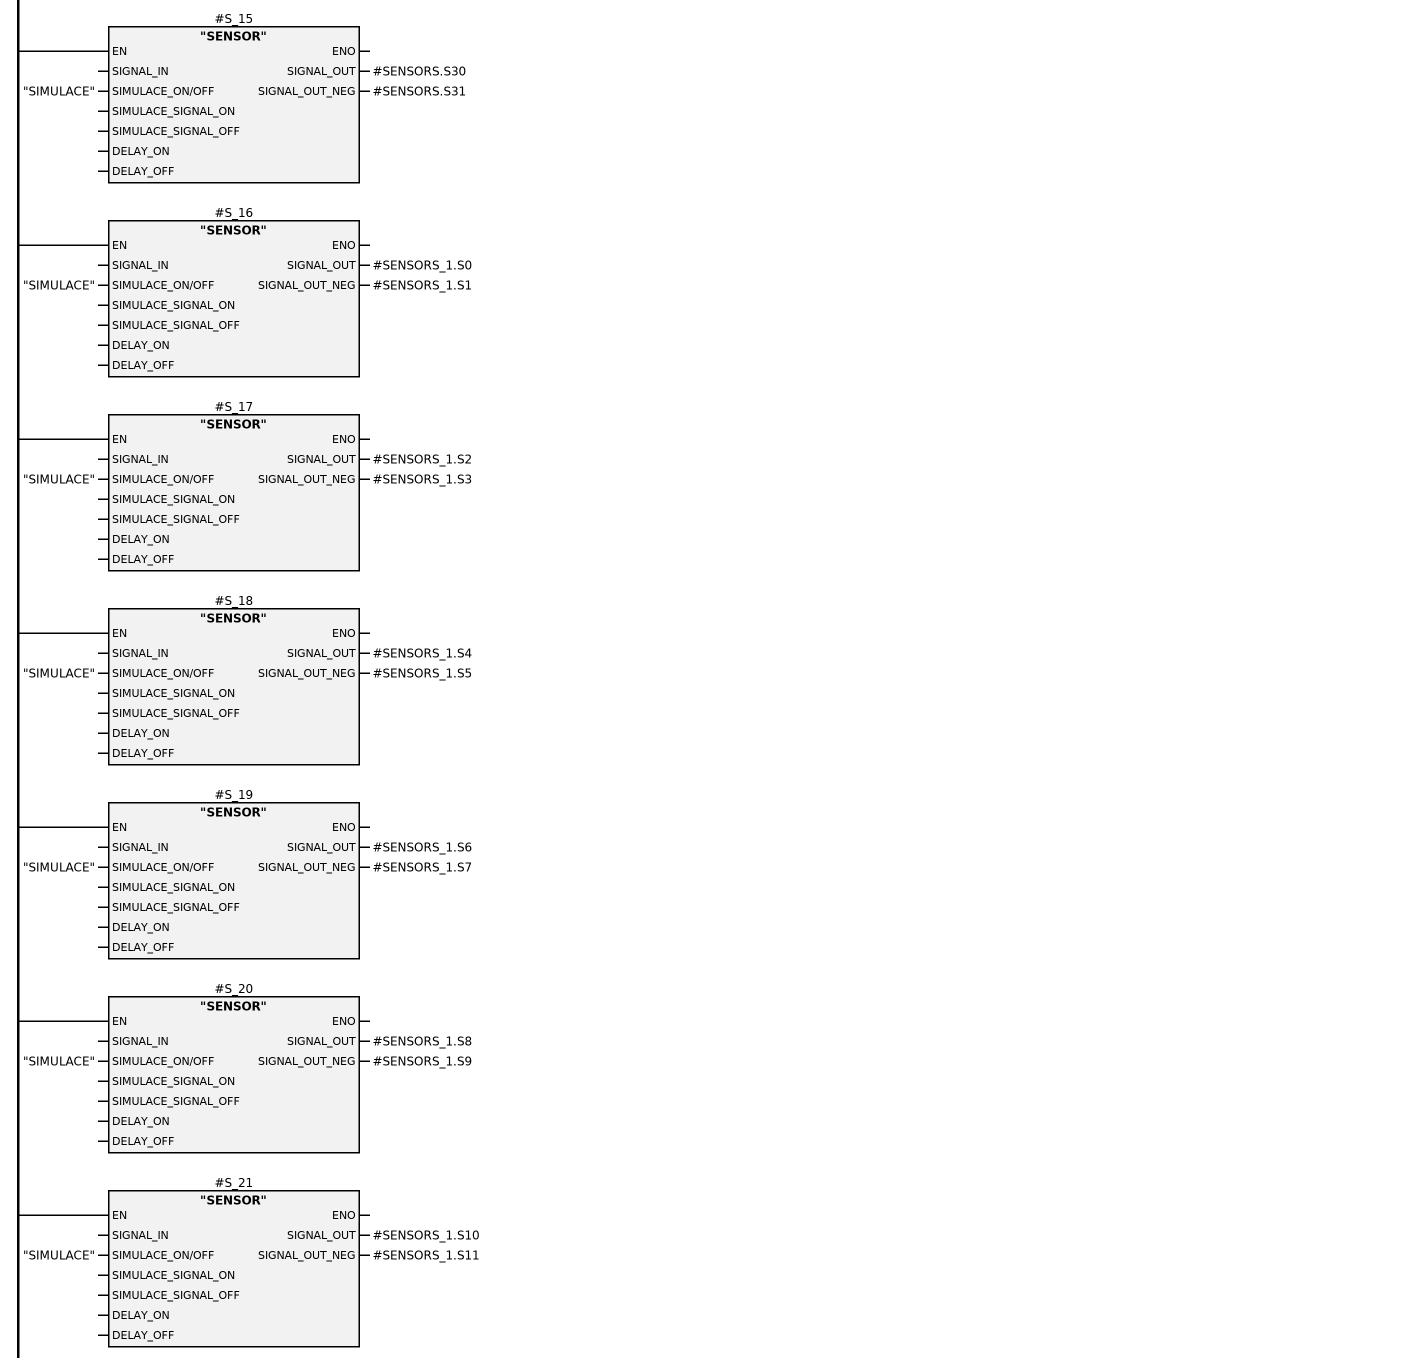
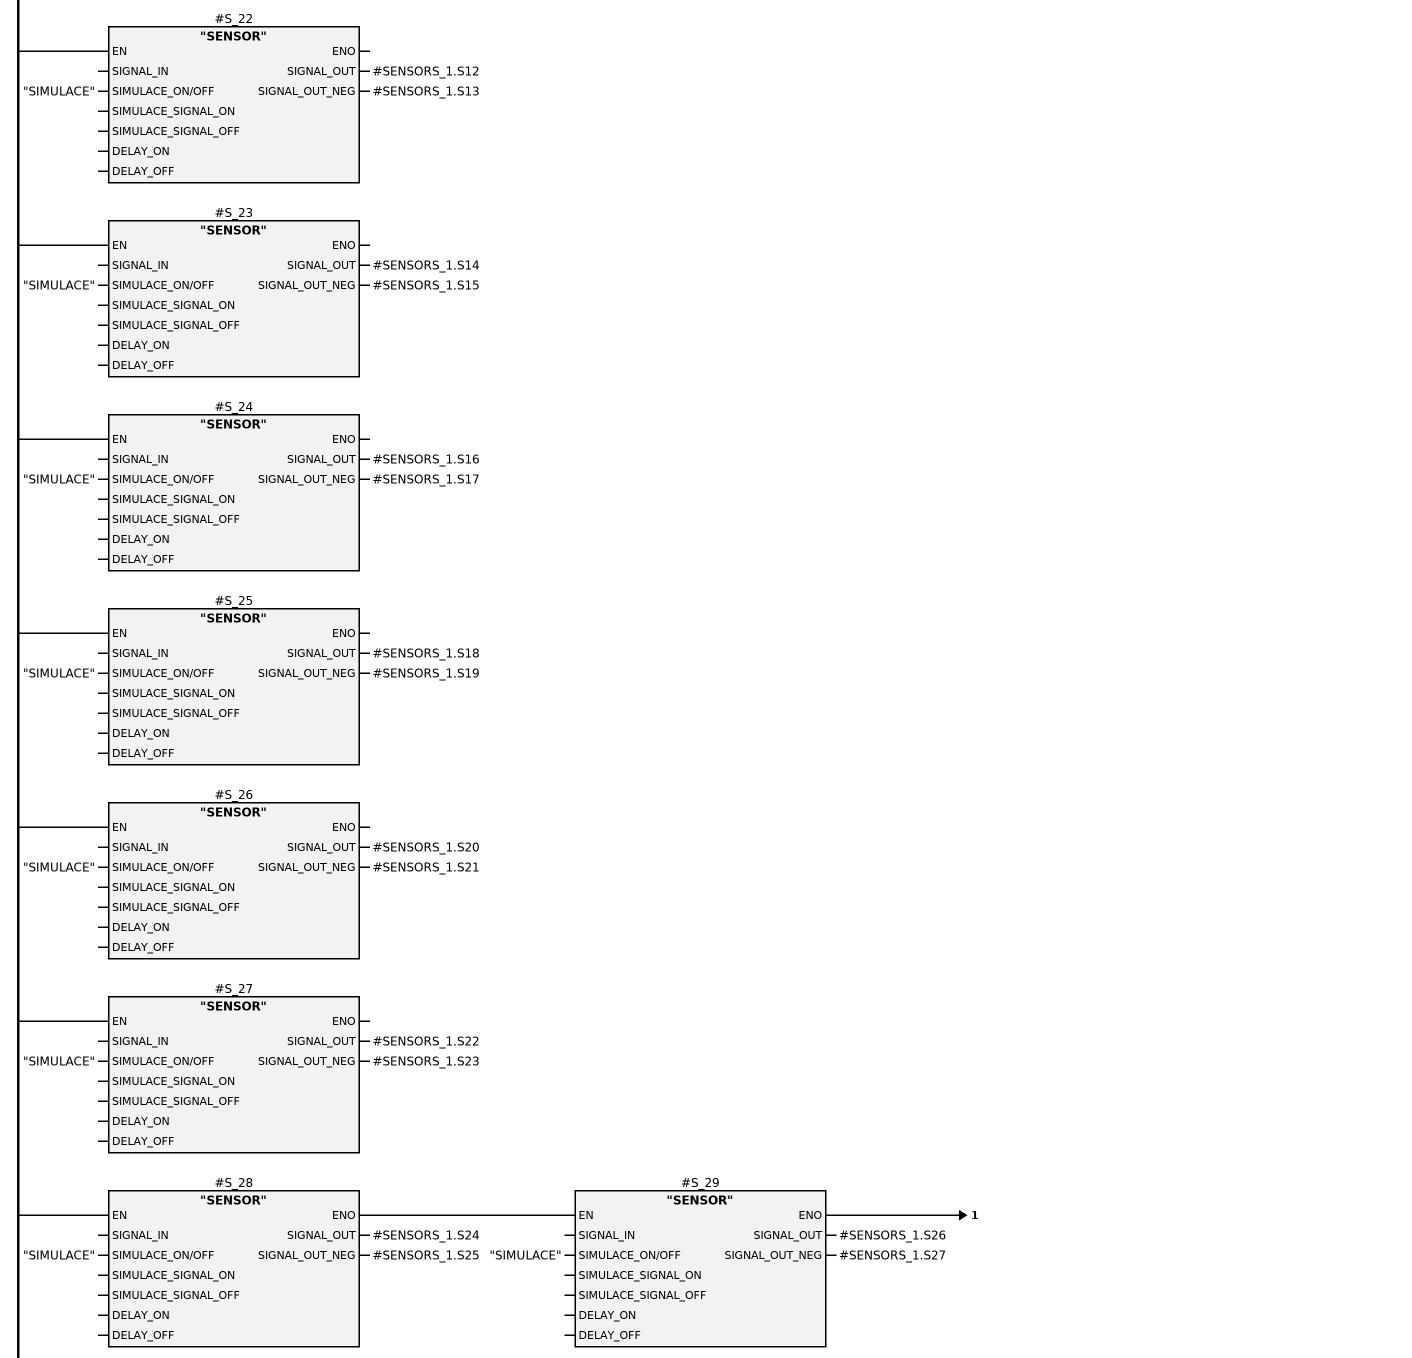
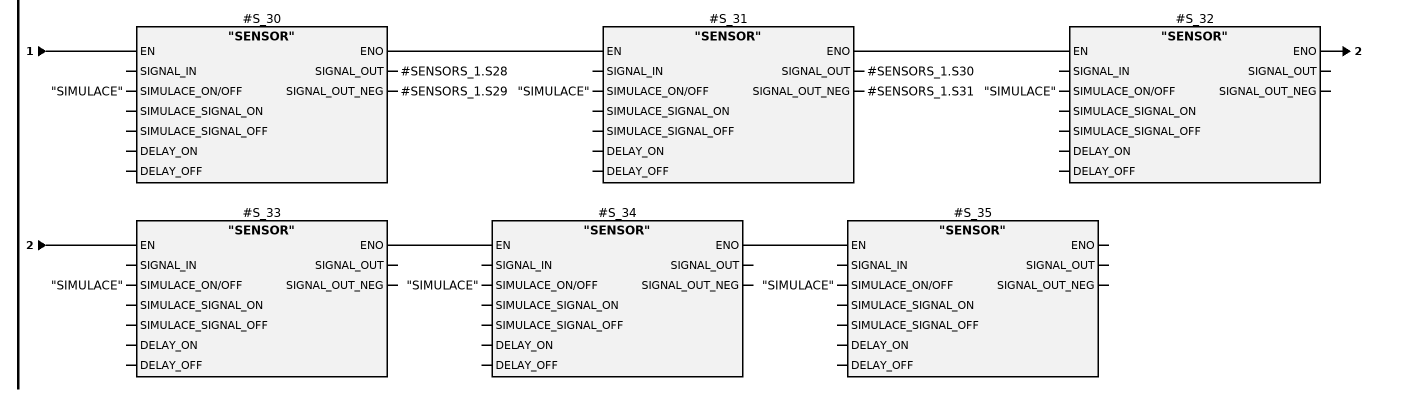
   RUNG wire#powerrail
      #S_0(SIGNAL_IN :=, "SIMULACE_ON/OFF" := "SIMULACE", SIMULACE_SIGNAL_ON :=, SIMULACE_SIGNAL_OFF :=, DELAY_ON :=, DELAY_OFF :=, SIGNAL_OUT => #SENSORS.S0, SIGNAL_OUT_NEG => #SENSORS.S1)
   END_RUNG
   RUNG wire#powerrail
      #S_1(SIGNAL_IN :=, "SIMULACE_ON/OFF" := "SIMULACE", SIMULACE_SIGNAL_ON :=, SIMULACE_SIGNAL_OFF :=, DELAY_ON :=, DELAY_OFF :=, SIGNAL_OUT => #SENSORS.S2, SIGNAL_OUT_NEG => #SENSORS.S3)
   END_RUNG
   RUNG wire#powerrail
      #S_2(SIGNAL_IN :=, "SIMULACE_ON/OFF" := "SIMULACE", SIMULACE_SIGNAL_ON :=, SIMULACE_SIGNAL_OFF :=, DELAY_ON :=, DELAY_OFF :=, SIGNAL_OUT => #SENSORS.S4, SIGNAL_OUT_NEG => #SENSORS.S5)
   END_RUNG
   RUNG wire#powerrail
      #S_3(SIGNAL_IN :=, "SIMULACE_ON/OFF" := "SIMULACE", SIMULACE_SIGNAL_ON :=, SIMULACE_SIGNAL_OFF :=, DELAY_ON :=, DELAY_OFF :=, SIGNAL_OUT => #SENSORS.S6, SIGNAL_OUT_NEG => #SENSORS.S7)
   END_RUNG
   RUNG wire#powerrail
      #S_4(SIGNAL_IN :=, "SIMULACE_ON/OFF" := "SIMULACE", SIMULACE_SIGNAL_ON :=, SIMULACE_SIGNAL_OFF :=, DELAY_ON :=, DELAY_OFF :=, SIGNAL_OUT => #SENSORS.S8, SIGNAL_OUT_NEG => #SENSORS.S9)
   END_RUNG
   RUNG wire#powerrail
      #S_6(SIGNAL_IN :=, "SIMULACE_ON/OFF" := "SIMULACE", SIMULACE_SIGNAL_ON :=, SIMULACE_SIGNAL_OFF :=, DELAY_ON :=, DELAY_OFF :=, SIGNAL_OUT => #SENSORS.S12, SIGNAL_OUT_NEG => #SENSORS.S13)
   END_RUNG
   RUNG wire#powerrail
      #S_5(SIGNAL_IN :=, "SIMULACE_ON/OFF" := "SIMULACE", SIMULACE_SIGNAL_ON :=, SIMULACE_SIGNAL_OFF :=, DELAY_ON :=, DELAY_OFF :=, SIGNAL_OUT => #SENSORS.S10, SIGNAL_OUT_NEG => #SENSORS.S11)
      #S_7(SIGNAL_IN :=, "SIMULACE_ON/OFF" := "SIMULACE", SIMULACE_SIGNAL_ON :=, SIMULACE_SIGNAL_OFF :=, DELAY_ON :=, DELAY_OFF :=, SIGNAL_OUT => #SENSORS.S14, SIGNAL_OUT_NEG => #SENSORS.S15)
      #S_8(SIGNAL_IN :=, "SIMULACE_ON/OFF" := "SIMULACE", SIMULACE_SIGNAL_ON :=, SIMULACE_SIGNAL_OFF :=, DELAY_ON :=, DELAY_OFF :=, SIGNAL_OUT => #SENSORS.S16, SIGNAL_OUT_NEG => #SENSORS.S17)
   END_RUNG
   RUNG wire#powerrail
      #S_9(SIGNAL_IN :=, "SIMULACE_ON/OFF" := "SIMULACE", SIMULACE_SIGNAL_ON :=, SIMULACE_SIGNAL_OFF :=, DELAY_ON :=, DELAY_OFF :=, SIGNAL_OUT => #SENSORS.S18, SIGNAL_OUT_NEG => #SENSORS.S19)
   END_RUNG
   RUNG wire#powerrail
      #s_10(SIGNAL_IN :=, "SIMULACE_ON/OFF" := "SIMULACE", SIMULACE_SIGNAL_ON :=, SIMULACE_SIGNAL_OFF :=, DELAY_ON :=, DELAY_OFF :=, SIGNAL_OUT => #SENSORS.S20, SIGNAL_OUT_NEG => #SENSORS.S21)
   END_RUNG
   RUNG wire#powerrail
      #S_11(SIGNAL_IN :=, "SIMULACE_ON/OFF" :=, SIMULACE_SIGNAL_ON := "SIMULACE", SIMULACE_SIGNAL_OFF :=, DELAY_ON :=, DELAY_OFF :=, SIGNAL_OUT => #SENSORS.S22, SIGNAL_OUT_NEG => #SENSORS.S23)
   END_RUNG
   RUNG wire#powerrail
      #S_12(SIGNAL_IN :=, "SIMULACE_ON/OFF" := "SIMULACE", SIMULACE_SIGNAL_ON :=, SIMULACE_SIGNAL_OFF :=, DELAY_ON :=, DELAY_OFF :=, SIGNAL_OUT => #SENSORS.S24, SIGNAL_OUT_NEG => #SENSORS.S25)
   END_RUNG
   RUNG wire#powerrail
      #S_13(SIGNAL_IN :=, "SIMULACE_ON/OFF" := "SIMULACE", SIMULACE_SIGNAL_ON :=, SIMULACE_SIGNAL_OFF :=, DELAY_ON :=, DELAY_OFF :=, SIGNAL_OUT => #SENSORS.S26, SIGNAL_OUT_NEG => #SENSORS.S27)
   END_RUNG
   RUNG wire#powerrail
      #S_14(SIGNAL_IN :=, "SIMULACE_ON/OFF" := "SIMULACE", SIMULACE_SIGNAL_ON :=, SIMULACE_SIGNAL_OFF :=, DELAY_ON :=, DELAY_OFF :=, SIGNAL_OUT => #SENSORS.S28, SIGNAL_OUT_NEG => #SENSORS.S29)
   END_RUNG
   RUNG wire#powerrail
      #S_15(SIGNAL_IN :=, "SIMULACE_ON/OFF" := "SIMULACE", SIMULACE_SIGNAL_ON :=, SIMULACE_SIGNAL_OFF :=, DELAY_ON :=, DELAY_OFF :=, SIGNAL_OUT => #SENSORS.S30, SIGNAL_OUT_NEG => #SENSORS.S31)
   END_RUNG
   RUNG wire#powerrail
      #S_16(SIGNAL_IN :=, "SIMULACE_ON/OFF" := "SIMULACE", SIMULACE_SIGNAL_ON :=, SIMULACE_SIGNAL_OFF :=, DELAY_ON :=, DELAY_OFF :=, SIGNAL_OUT => #SENSORS_1.S0, SIGNAL_OUT_NEG => #SENSORS_1.S1)
   END_RUNG
   RUNG wire#powerrail
      #S_17(SIGNAL_IN :=, "SIMULACE_ON/OFF" := "SIMULACE", SIMULACE_SIGNAL_ON :=, SIMULACE_SIGNAL_OFF :=, DELAY_ON :=, DELAY_OFF :=, SIGNAL_OUT => #SENSORS_1.S2, SIGNAL_OUT_NEG => #SENSORS_1.S3)
   END_RUNG
   RUNG wire#powerrail
      #S_18(SIGNAL_IN :=, "SIMULACE_ON/OFF" := "SIMULACE", SIMULACE_SIGNAL_ON :=, SIMULACE_SIGNAL_OFF :=, DELAY_ON :=, DELAY_OFF :=, SIGNAL_OUT => #SENSORS_1.S4, SIGNAL_OUT_NEG => #SENSORS_1.S5)
   END_RUNG
   RUNG wire#powerrail
      #S_19(SIGNAL_IN :=, "SIMULACE_ON/OFF" := "SIMULACE", SIMULACE_SIGNAL_ON :=, SIMULACE_SIGNAL_OFF :=, DELAY_ON :=, DELAY_OFF :=, SIGNAL_OUT => #SENSORS_1.S6, SIGNAL_OUT_NEG => #SENSORS_1.S7)
   END_RUNG
   RUNG wire#powerrail
      #S_20(SIGNAL_IN :=, "SIMULACE_ON/OFF" := "SIMULACE", SIMULACE_SIGNAL_ON :=, SIMULACE_SIGNAL_OFF :=, DELAY_ON :=, DELAY_OFF :=, SIGNAL_OUT => #SENSORS_1.S8, SIGNAL_OUT_NEG => #SENSORS_1.S9)
   END_RUNG
   RUNG wire#powerrail
      #S_21(SIGNAL_IN :=, "SIMULACE_ON/OFF" := "SIMULACE", SIMULACE_SIGNAL_ON :=, SIMULACE_SIGNAL_OFF :=, DELAY_ON :=, DELAY_OFF :=, SIGNAL_OUT => #SENSORS_1.S10, SIGNAL_OUT_NEG => #SENSORS_1.S11)
   END_RUNG
   RUNG wire#powerrail
      #S_22(SIGNAL_IN :=, "SIMULACE_ON/OFF" := "SIMULACE", SIMULACE_SIGNAL_ON :=, SIMULACE_SIGNAL_OFF :=, DELAY_ON :=, DELAY_OFF :=, SIGNAL_OUT => #SENSORS_1.S12, SIGNAL_OUT_NEG => #SENSORS_1.S13)
   END_RUNG
   RUNG wire#powerrail
      #S_23(SIGNAL_IN :=, "SIMULACE_ON/OFF" := "SIMULACE", SIMULACE_SIGNAL_ON :=, SIMULACE_SIGNAL_OFF :=, DELAY_ON :=, DELAY_OFF :=, SIGNAL_OUT => #SENSORS_1.S14, SIGNAL_OUT_NEG => #SENSORS_1.S15)
   END_RUNG
   RUNG wire#powerrail
      #S_24(SIGNAL_IN :=, "SIMULACE_ON/OFF" := "SIMULACE", SIMULACE_SIGNAL_ON :=, SIMULACE_SIGNAL_OFF :=, DELAY_ON :=, DELAY_OFF :=, SIGNAL_OUT => #SENSORS_1.S16, SIGNAL_OUT_NEG => #SENSORS_1.S17)
   END_RUNG
   RUNG wire#powerrail
      #S_25(SIGNAL_IN :=, "SIMULACE_ON/OFF" := "SIMULACE", SIMULACE_SIGNAL_ON :=, SIMULACE_SIGNAL_OFF :=, DELAY_ON :=, DELAY_OFF :=, SIGNAL_OUT => #SENSORS_1.S18, SIGNAL_OUT_NEG => #SENSORS_1.S19)
   END_RUNG
   RUNG wire#powerrail
      #S_26(SIGNAL_IN :=, "SIMULACE_ON/OFF" := "SIMULACE", SIMULACE_SIGNAL_ON :=, SIMULACE_SIGNAL_OFF :=, DELAY_ON :=, DELAY_OFF :=, SIGNAL_OUT => #SENSORS_1.S20, SIGNAL_OUT_NEG => #SENSORS_1.S21)
   END_RUNG
   RUNG wire#powerrail
      #S_27(SIGNAL_IN :=, "SIMULACE_ON/OFF" := "SIMULACE", SIMULACE_SIGNAL_ON :=, SIMULACE_SIGNAL_OFF :=, DELAY_ON :=, DELAY_OFF :=, SIGNAL_OUT => #SENSORS_1.S22, SIGNAL_OUT_NEG => #SENSORS_1.S23)
   END_RUNG
   RUNG wire#powerrail
      #S_28(SIGNAL_IN :=, "SIMULACE_ON/OFF" := "SIMULACE", SIMULACE_SIGNAL_ON :=, SIMULACE_SIGNAL_OFF :=, DELAY_ON :=, DELAY_OFF :=, SIGNAL_OUT => #SENSORS_1.S24, SIGNAL_OUT_NEG => #SENSORS_1.S25)
      #S_29(SIGNAL_IN :=, "SIMULACE_ON/OFF" := "SIMULACE", SIMULACE_SIGNAL_ON :=, SIMULACE_SIGNAL_OFF :=, DELAY_ON :=, DELAY_OFF :=, SIGNAL_OUT => #SENSORS_1.S26, SIGNAL_OUT_NEG => #SENSORS_1.S27)
      #S_30(SIGNAL_IN :=, "SIMULACE_ON/OFF" := "SIMULACE", SIMULACE_SIGNAL_ON :=, SIMULACE_SIGNAL_OFF :=, DELAY_ON :=, DELAY_OFF :=, SIGNAL_OUT => #SENSORS_1.S28, SIGNAL_OUT_NEG => #SENSORS_1.S29)
      #S_31(SIGNAL_IN :=, "SIMULACE_ON/OFF" := "SIMULACE", SIMULACE_SIGNAL_ON :=, SIMULACE_SIGNAL_OFF :=, DELAY_ON :=, DELAY_OFF :=, SIGNAL_OUT => #SENSORS_1.S30, SIGNAL_OUT_NEG => #SENSORS_1.S31)
      #S_32(SIGNAL_IN :=, "SIMULACE_ON/OFF" := "SIMULACE", SIMULACE_SIGNAL_ON :=, SIMULACE_SIGNAL_OFF :=, DELAY_ON :=, DELAY_OFF :=, SIGNAL_OUT =>, SIGNAL_OUT_NEG =>)
      #S_33(SIGNAL_IN :=, "SIMULACE_ON/OFF" := "SIMULACE", SIMULACE_SIGNAL_ON :=, SIMULACE_SIGNAL_OFF :=, DELAY_ON :=, DELAY_OFF :=, SIGNAL_OUT =>, SIGNAL_OUT_NEG =>)
      #S_34(SIGNAL_IN :=, "SIMULACE_ON/OFF" := "SIMULACE", SIMULACE_SIGNAL_ON :=, SIMULACE_SIGNAL_OFF :=, DELAY_ON :=, DELAY_OFF :=, SIGNAL_OUT =>, SIGNAL_OUT_NEG =>)
      #S_35(SIGNAL_IN :=, "SIMULACE_ON/OFF" := "SIMULACE", SIMULACE_SIGNAL_ON :=, SIMULACE_SIGNAL_OFF :=, DELAY_ON :=, DELAY_OFF :=, SIGNAL_OUT =>, SIGNAL_OUT_NEG =>)
   END_RUNG
   // the same network as SCL:
   #S_0("SIMULACE_ON/OFF" := "SIMULACE", SIGNAL_OUT => #SENSORS.S0, SIGNAL_OUT_NEG => #SENSORS.S1);   // "SENSOR"
   #S_1("SIMULACE_ON/OFF" := "SIMULACE", SIGNAL_OUT => #SENSORS.S2, SIGNAL_OUT_NEG => #SENSORS.S3);   // "SENSOR"
   #S_2("SIMULACE_ON/OFF" := "SIMULACE", SIGNAL_OUT => #SENSORS.S4, SIGNAL_OUT_NEG => #SENSORS.S5);   // "SENSOR"
   #S_3("SIMULACE_ON/OFF" := "SIMULACE", SIGNAL_OUT => #SENSORS.S6, SIGNAL_OUT_NEG => #SENSORS.S7);   // "SENSOR"
   #S_4("SIMULACE_ON/OFF" := "SIMULACE", SIGNAL_OUT => #SENSORS.S8, SIGNAL_OUT_NEG => #SENSORS.S9);   // "SENSOR"
   #S_6("SIMULACE_ON/OFF" := "SIMULACE", SIGNAL_OUT => #SENSORS.S12, SIGNAL_OUT_NEG => #SENSORS.S13);   // "SENSOR"
   #S_5("SIMULACE_ON/OFF" := "SIMULACE",   // "SENSOR"
        SIGNAL_OUT => #SENSORS.S10,
        SIGNAL_OUT_NEG => #SENSORS.S11,
        ENO => #_w1);
   #S_7(EN := #_w1,   // "SENSOR"
        "SIMULACE_ON/OFF" := "SIMULACE",
        SIGNAL_OUT => #SENSORS.S14,
        SIGNAL_OUT_NEG => #SENSORS.S15,
        ENO => #_w2);
   IF #_w2 THEN
       #S_8("SIMULACE_ON/OFF" := "SIMULACE", SIGNAL_OUT => #SENSORS.S16, SIGNAL_OUT_NEG => #SENSORS.S17);   // "SENSOR"
   END_IF;
   #S_9("SIMULACE_ON/OFF" := "SIMULACE", SIGNAL_OUT => #SENSORS.S18, SIGNAL_OUT_NEG => #SENSORS.S19);   // "SENSOR"
   #s_10("SIMULACE_ON/OFF" := "SIMULACE", SIGNAL_OUT => #SENSORS.S20, SIGNAL_OUT_NEG => #SENSORS.S21);   // "SENSOR"
   #S_11(SIMULACE_SIGNAL_ON := "SIMULACE", SIGNAL_OUT => #SENSORS.S22, SIGNAL_OUT_NEG => #SENSORS.S23);   // "SENSOR"
   #S_12("SIMULACE_ON/OFF" := "SIMULACE", SIGNAL_OUT => #SENSORS.S24, SIGNAL_OUT_NEG => #SENSORS.S25);   // "SENSOR"
   #S_13("SIMULACE_ON/OFF" := "SIMULACE", SIGNAL_OUT => #SENSORS.S26, SIGNAL_OUT_NEG => #SENSORS.S27);   // "SENSOR"
   #S_14("SIMULACE_ON/OFF" := "SIMULACE", SIGNAL_OUT => #SENSORS.S28, SIGNAL_OUT_NEG => #SENSORS.S29);   // "SENSOR"
   #S_15("SIMULACE_ON/OFF" := "SIMULACE", SIGNAL_OUT => #SENSORS.S30, SIGNAL_OUT_NEG => #SENSORS.S31);   // "SENSOR"
   #S_16("SIMULACE_ON/OFF" := "SIMULACE", SIGNAL_OUT => #SENSORS_1.S0, SIGNAL_OUT_NEG => #SENSORS_1.S1);   // "SENSOR"
   #S_17("SIMULACE_ON/OFF" := "SIMULACE", SIGNAL_OUT => #SENSORS_1.S2, SIGNAL_OUT_NEG => #SENSORS_1.S3);   // "SENSOR"
   #S_18("SIMULACE_ON/OFF" := "SIMULACE", SIGNAL_OUT => #SENSORS_1.S4, SIGNAL_OUT_NEG => #SENSORS_1.S5);   // "SENSOR"
   #S_19("SIMULACE_ON/OFF" := "SIMULACE", SIGNAL_OUT => #SENSORS_1.S6, SIGNAL_OUT_NEG => #SENSORS_1.S7);   // "SENSOR"
   #S_20("SIMULACE_ON/OFF" := "SIMULACE", SIGNAL_OUT => #SENSORS_1.S8, SIGNAL_OUT_NEG => #SENSORS_1.S9);   // "SENSOR"
   #S_21("SIMULACE_ON/OFF" := "SIMULACE", SIGNAL_OUT => #SENSORS_1.S10, SIGNAL_OUT_NEG => #SENSORS_1.S11);   // "SENSOR"
   #S_22("SIMULACE_ON/OFF" := "SIMULACE", SIGNAL_OUT => #SENSORS_1.S12, SIGNAL_OUT_NEG => #SENSORS_1.S13);   // "SENSOR"
   #S_23("SIMULACE_ON/OFF" := "SIMULACE", SIGNAL_OUT => #SENSORS_1.S14, SIGNAL_OUT_NEG => #SENSORS_1.S15);   // "SENSOR"
   #S_24("SIMULACE_ON/OFF" := "SIMULACE", SIGNAL_OUT => #SENSORS_1.S16, SIGNAL_OUT_NEG => #SENSORS_1.S17);   // "SENSOR"
   #S_25("SIMULACE_ON/OFF" := "SIMULACE", SIGNAL_OUT => #SENSORS_1.S18, SIGNAL_OUT_NEG => #SENSORS_1.S19);   // "SENSOR"
   #S_26("SIMULACE_ON/OFF" := "SIMULACE", SIGNAL_OUT => #SENSORS_1.S20, SIGNAL_OUT_NEG => #SENSORS_1.S21);   // "SENSOR"
   #S_27("SIMULACE_ON/OFF" := "SIMULACE", SIGNAL_OUT => #SENSORS_1.S22, SIGNAL_OUT_NEG => #SENSORS_1.S23);   // "SENSOR"
   #S_28("SIMULACE_ON/OFF" := "SIMULACE",   // "SENSOR"
         SIGNAL_OUT => #SENSORS_1.S24,
         SIGNAL_OUT_NEG => #SENSORS_1.S25,
         ENO => #_w3);
   #S_29(EN := #_w3,   // "SENSOR"
         "SIMULACE_ON/OFF" := "SIMULACE",
         SIGNAL_OUT => #SENSORS_1.S26,
         SIGNAL_OUT_NEG => #SENSORS_1.S27,
         ENO => #_w4);
   #S_30(EN := #_w4,   // "SENSOR"
         "SIMULACE_ON/OFF" := "SIMULACE",
         SIGNAL_OUT => #SENSORS_1.S28,
         SIGNAL_OUT_NEG => #SENSORS_1.S29,
         ENO => #_w5);
   #S_31(EN := #_w5,   // "SENSOR"
         "SIMULACE_ON/OFF" := "SIMULACE",
         SIGNAL_OUT => #SENSORS_1.S30,
         SIGNAL_OUT_NEG => #SENSORS_1.S31,
         ENO => #_w6);
   #S_32(EN := #_w6, "SIMULACE_ON/OFF" := "SIMULACE", ENO => #_w7);   // "SENSOR"
   #S_33(EN := #_w7, "SIMULACE_ON/OFF" := "SIMULACE", ENO => #_w8);   // "SENSOR"
   #S_34(EN := #_w8, "SIMULACE_ON/OFF" := "SIMULACE", ENO => #_w9);   // "SENSOR"
   IF #_w9 THEN
       #S_35("SIMULACE_ON/OFF" := "SIMULACE");   // "SENSOR"
   END_IF;
END_REGION

REGION Network 5: INICIALIZACE START
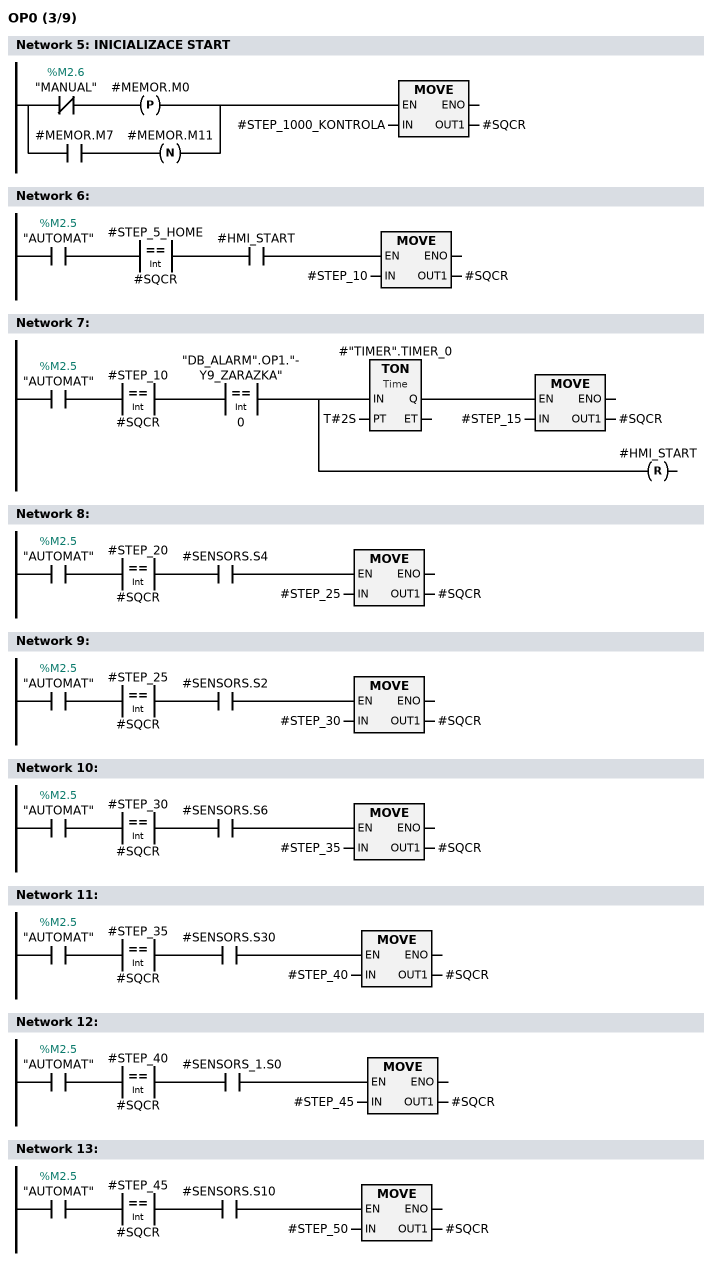
   RUNG wire#powerrail
      I_Contact( "MANUAL" )
      P_Trig( #MEMOR.M0 )
      wire#w1
      Move(in := #STEP_1000_KONTROLA, out1 => #SQCR)
   END_RUNG
   RUNG wire#powerrail
      Contact( #MEMOR.M7 )
      N_Trig( #MEMOR.M11 )
   END_RUNG wire#w1
   // the same network as SCL:
   #_w1 := NOT "MANUAL" AND NOT #MEMOR.M0;   // rising edge
   #MEMOR.M0 := NOT "MANUAL";
   #_w2 := NOT #MEMOR.M7 AND #MEMOR.M11;   // falling edge
   #MEMOR.M11 := #MEMOR.M7;
   IF #_w1 OR #_w2 THEN #SQCR := #STEP_1000_KONTROLA; END_IF;
END_REGION

REGION Network 6
   RUNG wire#powerrail
      Contact( "AUTOMAT" )
      { S7_Templates := "SrcType := Int" } EQ_Contact(in1 := #STEP_5_HOME, in2 := #SQCR)
      Contact( #HMI_START )
      Move(in := #STEP_10, out1 => #SQCR)
   END_RUNG
   // the same network as SCL:
   IF "AUTOMAT" AND (#STEP_5_HOME = #SQCR) AND #HMI_START THEN #SQCR := #STEP_10; END_IF;
END_REGION

REGION Network 7
   RUNG wire#powerrail
      Contact( "AUTOMAT" )
      { S7_Templates := "SrcType := Int" } EQ_Contact(in1 := #STEP_10, in2 := #SQCR)
      { S7_Templates := "SrcType := Int" } EQ_Contact(in1 := "DB_ALARM".OP1."-Y9_ZARAZKA", in2 := 0)
      wire#w1
      { S7_Templates := "time_type := Time" } #"TIMER".TIMER_0.TON(pt := T#2S, et =>)
      Move(in := #STEP_15, out1 => #SQCR)
   END_RUNG
   RUNG wire#w1
      R_Coil( #HMI_START )
   END_RUNG
   // the same network as SCL:
   #_w1 := "AUTOMAT" AND (#STEP_10 = #SQCR) AND ("DB_ALARM".OP1."-Y9_ZARAZKA" = 0);
   #"TIMER".TIMER_0.TON(IN := #_w1, PT := T#2S);
   IF #"TIMER".TIMER_0.Q THEN #SQCR := #STEP_15; END_IF;
   IF #_w1 THEN #HMI_START := FALSE; END_IF;
END_REGION

REGION Network 8
   RUNG wire#powerrail
      Contact( "AUTOMAT" )
      { S7_Templates := "SrcType := Int" } EQ_Contact(in1 := #STEP_20, in2 := #SQCR)
      Contact( #SENSORS.S4 )
      Move(in := #STEP_25, out1 => #SQCR)
   END_RUNG
   // the same network as SCL:
   IF "AUTOMAT" AND (#STEP_20 = #SQCR) AND #SENSORS.S4 THEN #SQCR := #STEP_25; END_IF;
END_REGION

REGION Network 9
   RUNG wire#powerrail
      Contact( "AUTOMAT" )
      { S7_Templates := "SrcType := Int" } EQ_Contact(in1 := #STEP_25, in2 := #SQCR)
      Contact( #SENSORS.S2 )
      Move(in := #STEP_30, out1 => #SQCR)
   END_RUNG
   // the same network as SCL:
   IF "AUTOMAT" AND (#STEP_25 = #SQCR) AND #SENSORS.S2 THEN #SQCR := #STEP_30; END_IF;
END_REGION

REGION Network 10
   RUNG wire#powerrail
      Contact( "AUTOMAT" )
      { S7_Templates := "SrcType := Int" } EQ_Contact(in1 := #STEP_30, in2 := #SQCR)
      Contact( #SENSORS.S6 )
      Move(in := #STEP_35, out1 => #SQCR)
   END_RUNG
   // the same network as SCL:
   IF "AUTOMAT" AND (#STEP_30 = #SQCR) AND #SENSORS.S6 THEN #SQCR := #STEP_35; END_IF;
END_REGION

REGION Network 11
   RUNG wire#powerrail
      Contact( "AUTOMAT" )
      { S7_Templates := "SrcType := Int" } EQ_Contact(in1 := #STEP_35, in2 := #SQCR)
      Contact( #SENSORS.S30 )
      Move(in := #STEP_40, out1 => #SQCR)
   END_RUNG
   // the same network as SCL:
   IF "AUTOMAT" AND (#STEP_35 = #SQCR) AND #SENSORS.S30 THEN #SQCR := #STEP_40; END_IF;
END_REGION

REGION Network 12
   RUNG wire#powerrail
      Contact( "AUTOMAT" )
      { S7_Templates := "SrcType := Int" } EQ_Contact(in1 := #STEP_40, in2 := #SQCR)
      Contact( #SENSORS_1.S0 )
      Move(in := #STEP_45, out1 => #SQCR)
   END_RUNG
   // the same network as SCL:
   IF "AUTOMAT" AND (#STEP_40 = #SQCR) AND #SENSORS_1.S0 THEN #SQCR := #STEP_45; END_IF;
END_REGION

REGION Network 13
   RUNG wire#powerrail
      Contact( "AUTOMAT" )
      { S7_Templates := "SrcType := Int" } EQ_Contact(in1 := #STEP_45, in2 := #SQCR)
      Contact( #SENSORS.S10 )
      Move(in := #STEP_50, out1 => #SQCR)
   END_RUNG
   // the same network as SCL:
   IF "AUTOMAT" AND (#STEP_45 = #SQCR) AND #SENSORS.S10 THEN #SQCR := #STEP_50; END_IF;
END_REGION

REGION Network 14
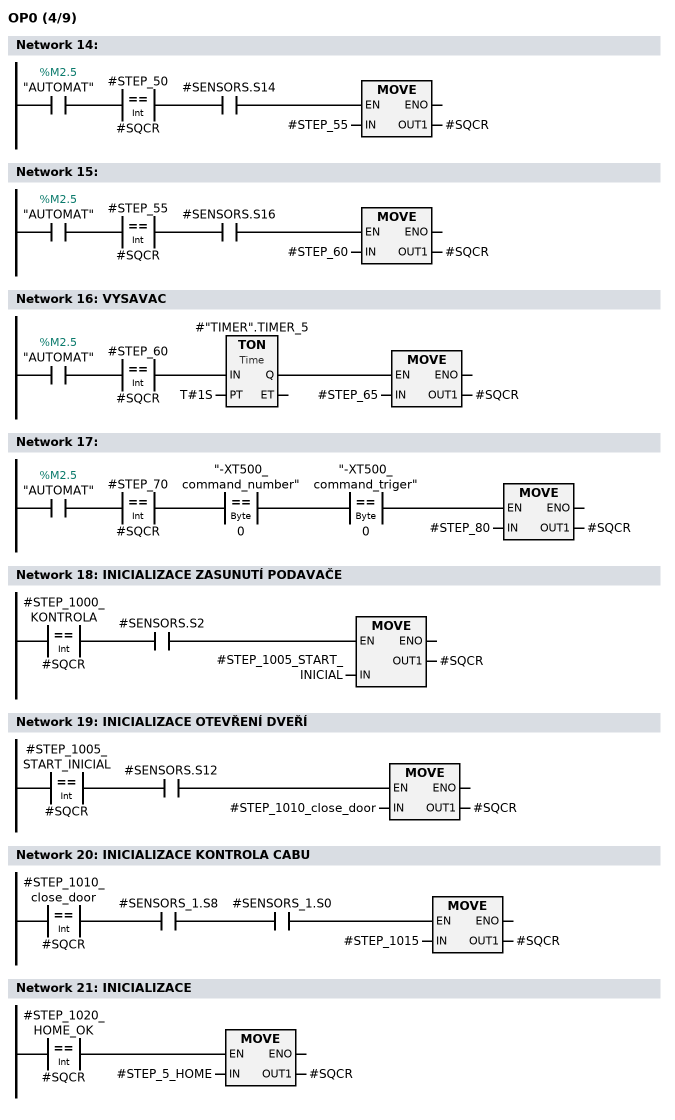
   RUNG wire#powerrail
      Contact( "AUTOMAT" )
      { S7_Templates := "SrcType := Int" } EQ_Contact(in1 := #STEP_50, in2 := #SQCR)
      Contact( #SENSORS.S14 )
      Move(in := #STEP_55, out1 => #SQCR)
   END_RUNG
   // the same network as SCL:
   IF "AUTOMAT" AND (#STEP_50 = #SQCR) AND #SENSORS.S14 THEN #SQCR := #STEP_55; END_IF;
END_REGION

REGION Network 15
   RUNG wire#powerrail
      Contact( "AUTOMAT" )
      { S7_Templates := "SrcType := Int" } EQ_Contact(in1 := #STEP_55, in2 := #SQCR)
      Contact( #SENSORS.S16 )
      Move(in := #STEP_60, out1 => #SQCR)
   END_RUNG
   // the same network as SCL:
   IF "AUTOMAT" AND (#STEP_55 = #SQCR) AND #SENSORS.S16 THEN #SQCR := #STEP_60; END_IF;
END_REGION

REGION Network 16: VYSAVAC
   RUNG wire#powerrail
      Contact( "AUTOMAT" )
      { S7_Templates := "SrcType := Int" } EQ_Contact(in1 := #STEP_60, in2 := #SQCR)
      { S7_Templates := "time_type := Time" } #"TIMER".TIMER_5.TON(pt := T#1S, et =>)
      Move(in := #STEP_65, out1 => #SQCR)
   END_RUNG
   // the same network as SCL:
   #"TIMER".TIMER_5.TON(IN := "AUTOMAT" AND (#STEP_60 = #SQCR), PT := T#1S);
   IF #"TIMER".TIMER_5.Q THEN #SQCR := #STEP_65; END_IF;
END_REGION

REGION Network 17
   RUNG wire#powerrail
      Contact( "AUTOMAT" )
      { S7_Templates := "SrcType := Int" } EQ_Contact(in1 := #STEP_70, in2 := #SQCR)
      { S7_Templates := "SrcType := Byte" } EQ_Contact(in1 := "-XT500_command_number", in2 := 0)
      { S7_Templates := "SrcType := Byte" } EQ_Contact(in1 := "-XT500_command_triger", in2 := 0)
      Move(in := #STEP_80, out1 => #SQCR)
   END_RUNG
   // the same network as SCL:
   IF "AUTOMAT" AND (#STEP_70 = #SQCR) AND ("-XT500_command_number" = 0) AND ("-XT500_command_triger" = 0) THEN
       #SQCR := #STEP_80;
   END_IF;
END_REGION

REGION Network 18: INICIALIZACE ZASUNUTÍ PODAVAČE
   RUNG wire#powerrail
      { S7_Templates := "SrcType := Int" } EQ_Contact(in1 := #STEP_1000_KONTROLA, in2 := #SQCR)
      Contact( #SENSORS.S2 )
      Move(in := #STEP_1005_START_INICIAL, out1 => #SQCR)
   END_RUNG
   // the same network as SCL:
   IF (#STEP_1000_KONTROLA = #SQCR) AND #SENSORS.S2 THEN #SQCR := #STEP_1005_START_INICIAL; END_IF;
END_REGION

REGION Network 19: INICIALIZACE OTEVŘENÍ DVEŘÍ
   RUNG wire#powerrail
      { S7_Templates := "SrcType := Int" } EQ_Contact(in1 := #STEP_1005_START_INICIAL, in2 := #SQCR)
      Contact( #SENSORS.S12 )
      Move(in := #STEP_1010_close_door, out1 => #SQCR)
   END_RUNG
   // the same network as SCL:
   IF (#STEP_1005_START_INICIAL = #SQCR) AND #SENSORS.S12 THEN #SQCR := #STEP_1010_close_door; END_IF;
END_REGION

REGION Network 20: INICIALIZACE KONTROLA CABU
   RUNG wire#powerrail
      { S7_Templates := "SrcType := Int" } EQ_Contact(in1 := #STEP_1010_close_door, in2 := #SQCR)
      Contact( #SENSORS_1.S8 )
      Contact( #SENSORS_1.S0 )
      Move(in := #STEP_1015, out1 => #SQCR)
   END_RUNG
   // the same network as SCL:
   IF (#STEP_1010_close_door = #SQCR) AND #SENSORS_1.S8 AND #SENSORS_1.S0 THEN #SQCR := #STEP_1015; END_IF;
END_REGION

REGION Network 21: INICIALIZACE
   RUNG wire#powerrail
      { S7_Templates := "SrcType := Int" } EQ_Contact(in1 := #STEP_1020_HOME_OK, in2 := #SQCR)
      Move(in := #STEP_5_HOME, out1 => #SQCR)
   END_RUNG
   // the same network as SCL:
   IF #STEP_1020_HOME_OK = #SQCR THEN #SQCR := #STEP_5_HOME; END_IF;
END_REGION

REGION Network 22: automat control door / automat control PODAVAC
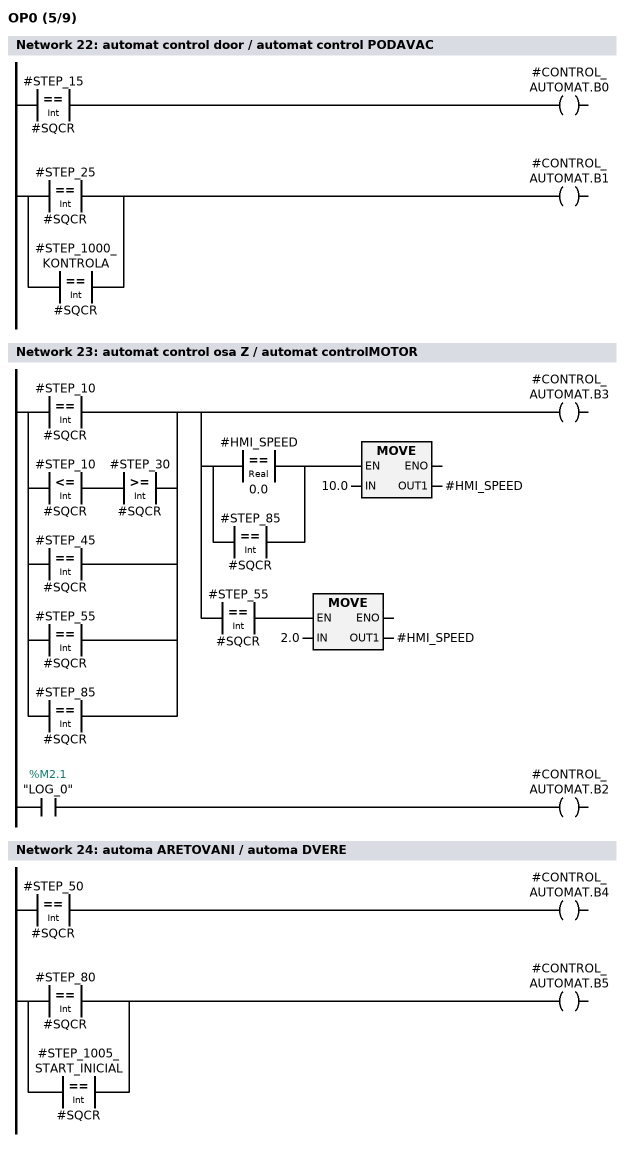
   RUNG wire#powerrail
      { S7_Templates := "SrcType := Int" } EQ_Contact(in1 := #STEP_15, in2 := #SQCR)
      Coil( #CONTROL_AUTOMAT.B0 )
   END_RUNG
   RUNG wire#powerrail
      { S7_Templates := "SrcType := Int" } EQ_Contact(in1 := #STEP_25, in2 := #SQCR)
      wire#w1
      Coil( #CONTROL_AUTOMAT.B1 )
   END_RUNG
   RUNG wire#powerrail
      { S7_Templates := "SrcType := Int" } EQ_Contact(in1 := #STEP_1000_KONTROLA, in2 := #SQCR)
   END_RUNG wire#w1
   // the same network as SCL:
   #CONTROL_AUTOMAT.B0 := #STEP_15 = #SQCR;
   #CONTROL_AUTOMAT.B1 := (#STEP_25 = #SQCR) OR (#STEP_1000_KONTROLA = #SQCR);
END_REGION

REGION Network 23: automat control osa Z / automat controlMOTOR
   RUNG wire#powerrail
      { S7_Templates := "SrcType := Int" } EQ_Contact(in1 := #STEP_10, in2 := #SQCR)
      wire#w1
      Coil( #CONTROL_AUTOMAT.B3 )
   END_RUNG
   RUNG wire#powerrail
      { S7_Templates := "SrcType := Int" } LE_Contact(in1 := #STEP_10, in2 := #SQCR)
      { S7_Templates := "SrcType := Int" } GE_Contact(in1 := #STEP_30, in2 := #SQCR)
   END_RUNG wire#w1
   RUNG wire#powerrail
      { S7_Templates := "SrcType := Int" } EQ_Contact(in1 := #STEP_45, in2 := #SQCR)
   END_RUNG wire#w1
   RUNG wire#powerrail
      { S7_Templates := "SrcType := Int" } EQ_Contact(in1 := #STEP_55, in2 := #SQCR)
   END_RUNG wire#w1
   RUNG wire#powerrail
      { S7_Templates := "SrcType := Int" } EQ_Contact(in1 := #STEP_85, in2 := #SQCR)
   END_RUNG wire#w1
   RUNG wire#w1
      { S7_Templates := "SrcType := Real" } EQ_Contact(in1 := #HMI_SPEED, in2 := 0.0)
      wire#w2
      Move(in := 10.0, out1 => #HMI_SPEED)
   END_RUNG
   RUNG wire#w1
      { S7_Templates := "SrcType := Int" } EQ_Contact(in1 := #STEP_85, in2 := #SQCR)
   END_RUNG wire#w2
   RUNG wire#w1
      { S7_Templates := "SrcType := Int" } EQ_Contact(in1 := #STEP_55, in2 := #SQCR)
      Move(in := 2.0, out1 => #HMI_SPEED)
   END_RUNG
   RUNG wire#powerrail
      Contact( "LOG_0" )
      Coil( #CONTROL_AUTOMAT.B2 )
   END_RUNG
   // the same network as SCL:
   #CONTROL_AUTOMAT.B3 := (#STEP_10 = #SQCR) OR ((#STEP_10 <= #SQCR) AND (#STEP_30 >= #SQCR)) OR (#STEP_45 = #SQCR) OR (#STEP_55 = #SQCR) OR (#STEP_85 = #SQCR);
   IF #CONTROL_AUTOMAT.B3 AND ((#HMI_SPEED = 0.0) OR (#STEP_85 = #SQCR)) THEN #HMI_SPEED := 10.0; END_IF;
   IF #CONTROL_AUTOMAT.B3 AND (#STEP_55 = #SQCR) THEN #HMI_SPEED := 2.0; END_IF;
   #CONTROL_AUTOMAT.B2 := "LOG_0";
END_REGION

REGION Network 24: automa ARETOVANI / automa DVERE
   RUNG wire#powerrail
      { S7_Templates := "SrcType := Int" } EQ_Contact(in1 := #STEP_50, in2 := #SQCR)
      Coil( #CONTROL_AUTOMAT.B4 )
   END_RUNG
   RUNG wire#powerrail
      { S7_Templates := "SrcType := Int" } EQ_Contact(in1 := #STEP_80, in2 := #SQCR)
      wire#w1
      Coil( #CONTROL_AUTOMAT.B5 )
   END_RUNG
   RUNG wire#powerrail
      { S7_Templates := "SrcType := Int" } EQ_Contact(in1 := #STEP_1005_START_INICIAL, in2 := #SQCR)
   END_RUNG wire#w1
   // the same network as SCL:
   #CONTROL_AUTOMAT.B4 := #STEP_50 = #SQCR;
   #CONTROL_AUTOMAT.B5 := (#STEP_80 = #SQCR) OR (#STEP_1005_START_INICIAL = #SQCR);
END_REGION

REGION Network 25: CONTROL BLOCK DVERE / CONTROL BLOCK podavač
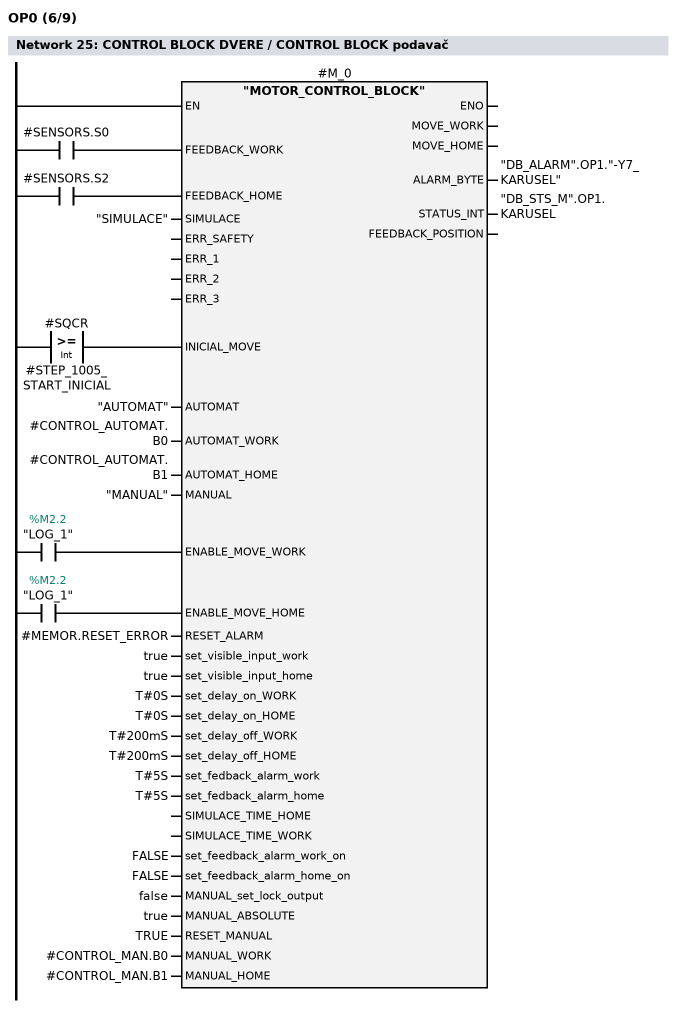
   RUNG wire#powerrail
      #M_0(FEEDBACK_WORK := wire#w1, FEEDBACK_HOME := wire#w2, INICIAL_MOVE := wire#w3, ENABLE_MOVE_WORK := wire#w4, ENABLE_MOVE_HOME := wire#w5, SIMULACE := "SIMULACE", ERR_SAFETY :=, ERR_1 :=, ERR_2 :=, ERR_3 :=, AUTOMAT := "AUTOMAT", AUTOMAT_WORK := #CONTROL_AUTOMAT.B0, AUTOMAT_HOME := #CONTROL_AUTOMAT.B1, MANUAL := "MANUAL", RESET_ALARM := #MEMOR.RESET_ERROR, set_visible_input_work := true, set_visible_input_home := true, set_delay_on_WORK := T#0S, set_delay_on_HOME := T#0S, set_delay_off_WORK := T#200mS, set_delay_off_HOME := T#200mS, set_fedback_alarm_work := T#5S, set_fedback_alarm_home := T#5S, SIMULACE_TIME_HOME :=, SIMULACE_TIME_WORK :=, set_feedback_alarm_work_on := FALSE, set_feedback_alarm_home_on := FALSE, MANUAL_set_lock_output := false, MANUAL_ABSOLUTE := true, RESET_MANUAL := TRUE, MANUAL_WORK := #CONTROL_MAN.B0, MANUAL_HOME := #CONTROL_MAN.B1, MOVE_WORK =>, MOVE_HOME =>, ALARM_BYTE => "DB_ALARM".OP1."-Y7_KARUSEL", STATUS_INT => "DB_STS_M".OP1.KARUSEL, FEEDBACK_POSITION =>)
   END_RUNG
   RUNG wire#powerrail
      Contact( #SENSORS.S0 )
   END_RUNG wire#w1
   RUNG wire#powerrail
      Contact( #SENSORS.S2 )
   END_RUNG wire#w2
   RUNG wire#powerrail
      { S7_Templates := "SrcType := Int" } GE_Contact(in1 := #SQCR, in2 := #STEP_1005_START_INICIAL)
   END_RUNG wire#w3
   RUNG wire#powerrail
      Contact( "LOG_1" )
   END_RUNG wire#w4
   RUNG wire#powerrail
      Contact( "LOG_1" )
   END_RUNG wire#w5
   // the same network as SCL:
   #M_0(FEEDBACK_WORK := #SENSORS.S0,   // "MOTOR_CONTROL_BLOCK"
        FEEDBACK_HOME := #SENSORS.S2,
        SIMULACE := "SIMULACE",
        INICIAL_MOVE := #SQCR >= #STEP_1005_START_INICIAL,
        AUTOMAT := "AUTOMAT",
        AUTOMAT_WORK := #CONTROL_AUTOMAT.B0,
        AUTOMAT_HOME := #CONTROL_AUTOMAT.B1,
        MANUAL := "MANUAL",
        ENABLE_MOVE_WORK := "LOG_1",
        ENABLE_MOVE_HOME := "LOG_1",
        RESET_ALARM := #MEMOR.RESET_ERROR,
        set_visible_input_work := true,
        set_visible_input_home := true,
        set_delay_on_WORK := T#0S,
        set_delay_on_HOME := T#0S,
        set_delay_off_WORK := T#200mS,
        set_delay_off_HOME := T#200mS,
        set_fedback_alarm_work := T#5S,
        set_fedback_alarm_home := T#5S,
        set_feedback_alarm_work_on := FALSE,
        set_feedback_alarm_home_on := FALSE,
        MANUAL_set_lock_output := false,
        MANUAL_ABSOLUTE := true,
        RESET_MANUAL := TRUE,
        MANUAL_WORK := #CONTROL_MAN.B0,
        MANUAL_HOME := #CONTROL_MAN.B1,
        ALARM_BYTE => "DB_ALARM".OP1."-Y7_KARUSEL",
        STATUS_INT => "DB_STS_M".OP1.KARUSEL);
END_REGION

REGION Network 26: CONTROL BLOCK OSA Z / CONTROL BLOCK dopravník
